// ---- DUTs/IO/Topology/Device_4_EtherCAT_07442C6B.TcDUT
{attribute 'GeneratedUsingTerminal: IODEVICETYPE_ETHERCATPROT'}
{attribute addProperty BoxType "IODEVICETYPE_ETHERCATPROT"}
{attribute addProperty Id "R1_EK1100R1_EK1100_4AD22B7B1143R2_EK1100R2_EK1100_10D8A594458R3_EK1100R3_EK1100_C7887D6C263R4_EK1100R4_EK1100_46A1248C369R4A_EK1100R4A_EK1100_48316913274R5_EK1100R5_EK1100_0007A337146R6_EK1100R6_EK1100_8C41F5F2336R7_EK1100R7_EK1100_F50DDAC8306R8_EK1100R8_EK1100_9C7B3B675648R9_EK1100R9_EK1100_484053C0136R10_EK1100R10_EK1100_C5CE1D87649SyncUnitsSyncUnits_5BE71B8B288InputsInputs_A65FACA410OutputsOutputs_23C0ED1D6InfoDataInfoData_84133AC922"}
{attribute addProperty CRC "121908331"}
{attribute addProperty Size "10054"}
{attribute addProperty Name "Device 4 (EtherCAT)"}
TYPE Device_4_EtherCAT_07442C6B EXTENDS TcoIo.EtcMasterBase_62654B43 :
STRUCT
	{attribute addProperty Name "R1 (EK1100)"}
	{attribute addProperty PreviousPort "Device 4 (EtherCAT) : Master"}
	{attribute addProperty SyncUnit "default"}
	R1_EK1100 : R1_EK1100_4AD22B7B;
	{attribute addProperty Name "R2 (EK1100)"}
	{attribute addProperty PreviousPort "R1 (EK1100) : C"}
	{attribute addProperty SyncUnit "default"}
	R2_EK1100 : R2_EK1100_10D8A594;
	{attribute addProperty Name "R3 (EK1100)"}
	{attribute addProperty PreviousPort "R2 (EK1100) : C"}
	{attribute addProperty SyncUnit "default"}
	R3_EK1100 : R3_EK1100_C7887D6C;
	{attribute addProperty Name "R4 (EK1100)"}
	{attribute addProperty PreviousPort "R3 (EK1100) : C"}
	{attribute addProperty SyncUnit "default"}
	R4_EK1100 : R4_EK1100_46A1248C;
	{attribute addProperty Name "R4A (EK1100)"}
	{attribute addProperty PreviousPort "R4 (EK1100) : C"}
	{attribute addProperty SyncUnit "default"}
	R4A_EK1100 : R4A_EK1100_48316913;
	{attribute addProperty Name "R5 (EK1100)"}
	{attribute addProperty PreviousPort "R4A (EK1100) : C"}
	{attribute addProperty SyncUnit "default"}
	R5_EK1100 : R5_EK1100_0007A337;
	{attribute addProperty Name "R6 (EK1100)"}
	{attribute addProperty PreviousPort "R5 (EK1100) : C"}
	{attribute addProperty SyncUnit "default"}
	R6_EK1100 : R6_EK1100_8C41F5F2;
	{attribute addProperty Name "R7 (EK1100)"}
	{attribute addProperty PreviousPort "R6 (EK1100) : C"}
	{attribute addProperty SyncUnit "default"}
	R7_EK1100 : R7_EK1100_F50DDAC8;
	{attribute addProperty Name "R8 (EK1100)"}
	{attribute addProperty PreviousPort "R7 (EK1100) : C"}
	{attribute addProperty SyncUnit "default"}
	R8_EK1100 : R8_EK1100_9C7B3B67;
	{attribute addProperty Name "R9 (EK1100)"}
	{attribute addProperty PreviousPort "R8 (EK1100) : C"}
	{attribute addProperty SyncUnit "default"}
	R9_EK1100 : R9_EK1100_484053C0;
	{attribute addProperty Name "R10 (EK1100)"}
	{attribute addProperty PreviousPort "R9 (EK1100) : C"}
	{attribute addProperty SyncUnit "default"}
	R10_EK1100 : R10_EK1100_C5CE1D87;
	{attribute addProperty Name "SyncUnits"}
	SyncUnits : SyncUnits_5BE71B8B;
	{attribute addProperty Name "Inputs"}
	Inputs : TcoIo.Inputs_A65FACA4;
	{attribute addProperty Name "Outputs"}
	Outputs : TcoIo.Outputs_23C0ED1D;
	{attribute addProperty Name "InfoData"}
	InfoData : TcoIo.InfoData_84133AC9;
END_STRUCT
END_TYPE

// ---- DUTs/IO/Topology/Term_279_EK1100_ED7D6272.TcDUT
{attribute 'GeneratedUsingTerminal: EK1100-0000-0018'}
{attribute addProperty BoxType "EK1100-0000-0018"}
{attribute addProperty Id "Term_280_EL1809EL1809_32157CFD20Term_281_EL1809EL1809_32157CFD20Term_282_EL1809EL1809_32157CFD20Term_283_EL1809EL1809_32157CFD20Term_284_EL1809EL1809_32157CFD20Term_312_EL1809EL1809_32157CFD20Term_320_EL1809EL1809_32157CFD20Term_321_EL1809EL1809_32157CFD20Term_322_EL1809EL1809_32157CFD20Term_323_EL1809EL1809_32157CFD20Term_324_EL1809EL1809_32157CFD20Term_325_EL1809EL1809_32157CFD20Term_326_EL1809EL1809_32157CFD20Term_327_EL1809EL1809_32157CFD20Term_328_EL1809EL1809_32157CFD20Term_329_EL1809EL1809_32157CFD20Term_331_EL1809EL1809_32157CFD20Term_332_EL1809EL1809_32157CFD20Term_333_EL1809EL1809_32157CFD20Term_334_EL1809EL1809_32157CFD20Term_335_EL1809EL1809_32157CFD20Term_336_EL1809EL1809_32157CFD20Term_337_EL1809EL1809_32157CFD20Term_338_EL1809EL1809_32157CFD20Term_339_EL1809EL1809_32157CFD20Term_340_EL1809EL1809_32157CFD20Term_341_EL1809EL1809_32157CFD20Term_342_EL1809EL1809_32157CFD20Term_343_EL1809EL1809_32157CFD20Term_344_EL1809EL1809_32157CFD20Term_345_EL1809EL1809_32157CFD20Term_346_EL1809EL1809_32157CFD20Term_347_EL1809EL1809_32157CFD20Term_348_EL1809EL1809_32157CFD20Term_360_EL1809EL1809_32157CFD20Term_361_EL1809EL1809_32157CFD20Term_362_EL1809EL1809_32157CFD20Term_363_EL1809EL1809_32157CFD20Term_364_EL1809EL1809_32157CFD20Term_365_EL1809EL1809_32157CFD20Term_366_EL1809EL1809_32157CFD20Term_367_EL1809EL1809_32157CFD20Term_368_EL1809EL1809_32157CFD20Term_370_EL1809EL1809_32157CFD20Term_371_EL1809EL1809_32157CFD20Term_372_EL1809EL1809_32157CFD20Term_373_EL1809EL1809_32157CFD20Term_374_EL1809EL1809_32157CFD20Term_375_EL1809EL1809_32157CFD20Term_376_EL1809EL1809_32157CFD20Term_377_EL1809EL1809_32157CFD20Term_378_EL1809EL1809_32157CFD20Term_380_EL1809EL1809_32157CFD20Term_381_EL1809EL1809_32157CFD20Term_382_EL1809EL1809_32157CFD20Term_383_EL1809EL1809_32157CFD20Term_384_EL1809EL1809_32157CFD20Term_385_EL1809EL1809_32157CFD20Term_386_EL1809EL1809_32157CFD20Term_387_EL1809EL1809_32157CFD20Term_388_EL1809EL1809_32157CFD20Term_389_EL1809EL1809_32157CFD20Term_390_EL1809EL1809_32157CFD20Term_391_EL1809EL1809_32157CFD20Term_392_EL1809EL1809_32157CFD20Term_393_EL1809EL1809_32157CFD20Term_394_EL1809EL1809_32157CFD20Term_395_EL1809EL1809_32157CFD20Term_396_EL1809EL1809_32157CFD20Term_397_EL1809EL1809_32157CFD20Term_398_EL1809EL1809_32157CFD20Term_399_EL1809EL1809_32157CFD20Term_400_EL1809EL1809_32157CFD20Term_401_EL1809EL1809_32157CFD20Term_402_EL1809EL1809_32157CFD20Term_403_EL1809EL1809_32157CFD20Term_404_EL1809EL1809_32157CFD20Term_405_EL1809EL1809_32157CFD20Term_406_EL1809EL1809_32157CFD20Term_407_EL1809EL1809_32157CFD20Term_408_EL1809EL1809_32157CFD20Term_409_EL1809EL1809_32157CFD20Term_410_EL1809EL1809_32157CFD20Term_414_EL1809EL1809_32157CFD20Term_415_EL1809EL1809_32157CFD20Term_416_EL1809EL1809_32157CFD20Term_417_EL1809EL1809_32157CFD20Term_418_EL1809EL1809_32157CFD20Term_419_EL1809EL1809_32157CFD20Term_420_EL1809EL1809_32157CFD20Term_421_EL1809EL1809_32157CFD20Term_422_EL1809EL1809_32157CFD20Term_423_EL1809EL1809_32157CFD20Term_424_EL1809EL1809_32157CFD20Term_425_EL1809EL1809_32157CFD20Term_426_EL1809EL1809_32157CFD20Term_427_EL1809EL1809_32157CFD20Term_428_EL1809EL1809_32157CFD20Term_429_EL1809EL1809_32157CFD20Term_448_EL1809EL1809_32157CFD20Term_495_EK1110EK1110_1FC0878B2"}
{attribute addProperty CRC "3984417394"}
{attribute addProperty Size "2002"}
{attribute addProperty Name "Term 279 (EK1100)"}
TYPE Term_279_EK1100_ED7D6272 EXTENDS EK1100_1FC0878B :
STRUCT
	{attribute addProperty Name "Term 280 (EL1809)"}
	{attribute addProperty PreviousPort "Term 279 (EK1100) : B"}
	{attribute addProperty SyncUnit "default"}
	Term_280_EL1809 : EL1809_32157CFD;
	{attribute addProperty Name "Term 281 (EL1809)"}
	{attribute addProperty PreviousPort "Term 280 (EL1809) : B"}
	{attribute addProperty SyncUnit "default"}
	Term_281_EL1809 : EL1809_32157CFD;
	{attribute addProperty Name "Term 282 (EL1809)"}
	{attribute addProperty PreviousPort "Term 281 (EL1809) : B"}
	{attribute addProperty SyncUnit "default"}
	Term_282_EL1809 : EL1809_32157CFD;
	{attribute addProperty Name "Term 283 (EL1809)"}
	{attribute addProperty PreviousPort "Term 282 (EL1809) : B"}
	{attribute addProperty SyncUnit "default"}
	Term_283_EL1809 : EL1809_32157CFD;
	{attribute addProperty Name "Term 284 (EL1809)"}
	{attribute addProperty PreviousPort "Term 283 (EL1809) : B"}
	{attribute addProperty SyncUnit "default"}
	Term_284_EL1809 : EL1809_32157CFD;
	{attribute addProperty Name "Term 312 (EL1809)"}
	{attribute addProperty PreviousPort "Term 284 (EL1809) : B"}
	{attribute addProperty SyncUnit "default"}
	Term_312_EL1809 : EL1809_32157CFD;
	{attribute addProperty Name "Term 320 (EL1809)"}
	{attribute addProperty PreviousPort "Term 312 (EL1809) : B"}
	{attribute addProperty SyncUnit "default"}
	Term_320_EL1809 : EL1809_32157CFD;
	{attribute addProperty Name "Term 321 (EL1809)"}
	{attribute addProperty PreviousPort "Term 320 (EL1809) : B"}
	{attribute addProperty SyncUnit "default"}
	Term_321_EL1809 : EL1809_32157CFD;
	{attribute addProperty Name "Term 322 (EL1809)"}
	{attribute addProperty PreviousPort "Term 321 (EL1809) : B"}
	{attribute addProperty SyncUnit "default"}
	Term_322_EL1809 : EL1809_32157CFD;
	{attribute addProperty Name "Term 323 (EL1809)"}
	{attribute addProperty PreviousPort "Term 322 (EL1809) : B"}
	{attribute addProperty SyncUnit "default"}
	Term_323_EL1809 : EL1809_32157CFD;
	{attribute addProperty Name "Term 324 (EL1809)"}
	{attribute addProperty PreviousPort "Term 323 (EL1809) : B"}
	{attribute addProperty SyncUnit "default"}
	Term_324_EL1809 : EL1809_32157CFD;
	{attribute addProperty Name "Term 325 (EL1809)"}
	{attribute addProperty PreviousPort "Term 324 (EL1809) : B"}
	{attribute addProperty SyncUnit "default"}
	Term_325_EL1809 : EL1809_32157CFD;
	{attribute addProperty Name "Term 326 (EL1809)"}
	{attribute addProperty PreviousPort "Term 325 (EL1809) : B"}
	{attribute addProperty SyncUnit "default"}
	Term_326_EL1809 : EL1809_32157CFD;
	{attribute addProperty Name "Term 327 (EL1809)"}
	{attribute addProperty PreviousPort "Term 326 (EL1809) : B"}
	{attribute addProperty SyncUnit "default"}
	Term_327_EL1809 : EL1809_32157CFD;
	{attribute addProperty Name "Term 328 (EL1809)"}
	{attribute addProperty PreviousPort "Term 327 (EL1809) : B"}
	{attribute addProperty SyncUnit "default"}
	Term_328_EL1809 : EL1809_32157CFD;
	{attribute addProperty Name "Term 329 (EL1809)"}
	{attribute addProperty PreviousPort "Term 328 (EL1809) : B"}
	{attribute addProperty SyncUnit "default"}
	Term_329_EL1809 : EL1809_32157CFD;
	{attribute addProperty Name "Term 331 (EL1809)"}
	{attribute addProperty PreviousPort "Term 329 (EL1809) : B"}
	{attribute addProperty SyncUnit "default"}
	Term_331_EL1809 : EL1809_32157CFD;
	{attribute addProperty Name "Term 332 (EL1809)"}
	{attribute addProperty PreviousPort "Term 331 (EL1809) : B"}
	{attribute addProperty SyncUnit "default"}
	Term_332_EL1809 : EL1809_32157CFD;
	{attribute addProperty Name "Term 333 (EL1809)"}
	{attribute addProperty PreviousPort "Term 332 (EL1809) : B"}
	{attribute addProperty SyncUnit "default"}
	Term_333_EL1809 : EL1809_32157CFD;
	{attribute addProperty Name "Term 334 (EL1809)"}
	{attribute addProperty PreviousPort "Term 333 (EL1809) : B"}
	{attribute addProperty SyncUnit "default"}
	Term_334_EL1809 : EL1809_32157CFD;
	{attribute addProperty Name "Term 335 (EL1809)"}
	{attribute addProperty PreviousPort "Term 334 (EL1809) : B"}
	{attribute addProperty SyncUnit "default"}
	Term_335_EL1809 : EL1809_32157CFD;
	{attribute addProperty Name "Term 336 (EL1809)"}
	{attribute addProperty PreviousPort "Term 335 (EL1809) : B"}
	{attribute addProperty SyncUnit "default"}
	Term_336_EL1809 : EL1809_32157CFD;
	{attribute addProperty Name "Term 337 (EL1809)"}
	{attribute addProperty PreviousPort "Term 336 (EL1809) : B"}
	{attribute addProperty SyncUnit "default"}
	Term_337_EL1809 : EL1809_32157CFD;
	{attribute addProperty Name "Term 338 (EL1809)"}
	{attribute addProperty PreviousPort "Term 337 (EL1809) : B"}
	{attribute addProperty SyncUnit "default"}
	Term_338_EL1809 : EL1809_32157CFD;
	{attribute addProperty Name "Term 339 (EL1809)"}
	{attribute addProperty PreviousPort "Term 338 (EL1809) : B"}
	{attribute addProperty SyncUnit "default"}
	Term_339_EL1809 : EL1809_32157CFD;
	{attribute addProperty Name "Term 340 (EL1809)"}
	{attribute addProperty PreviousPort "Term 339 (EL1809) : B"}
	{attribute addProperty SyncUnit "default"}
	Term_340_EL1809 : EL1809_32157CFD;
	{attribute addProperty Name "Term 341 (EL1809)"}
	{attribute addProperty PreviousPort "Term 340 (EL1809) : B"}
	{attribute addProperty SyncUnit "default"}
	Term_341_EL1809 : EL1809_32157CFD;
	{attribute addProperty Name "Term 342 (EL1809)"}
	{attribute addProperty PreviousPort "Term 341 (EL1809) : B"}
	{attribute addProperty SyncUnit "default"}
	Term_342_EL1809 : EL1809_32157CFD;
	{attribute addProperty Name "Term 343 (EL1809)"}
	{attribute addProperty PreviousPort "Term 342 (EL1809) : B"}
	{attribute addProperty SyncUnit "default"}
	Term_343_EL1809 : EL1809_32157CFD;
	{attribute addProperty Name "Term 344 (EL1809)"}
	{attribute addProperty PreviousPort "Term 343 (EL1809) : B"}
	{attribute addProperty SyncUnit "default"}
	Term_344_EL1809 : EL1809_32157CFD;
	{attribute addProperty Name "Term 345 (EL1809)"}
	{attribute addProperty PreviousPort "Term 344 (EL1809) : B"}
	{attribute addProperty SyncUnit "default"}
	Term_345_EL1809 : EL1809_32157CFD;
	{attribute addProperty Name "Term 346 (EL1809)"}
	{attribute addProperty PreviousPort "Term 345 (EL1809) : B"}
	{attribute addProperty SyncUnit "default"}
	Term_346_EL1809 : EL1809_32157CFD;
	{attribute addProperty Name "Term 347 (EL1809)"}
	{attribute addProperty PreviousPort "Term 346 (EL1809) : B"}
	{attribute addProperty SyncUnit "default"}
	Term_347_EL1809 : EL1809_32157CFD;
	{attribute addProperty Name "Term 348 (EL1809)"}
	{attribute addProperty PreviousPort "Term 347 (EL1809) : B"}
	{attribute addProperty SyncUnit "default"}
	Term_348_EL1809 : EL1809_32157CFD;
	{attribute addProperty Name "Term 360 (EL1809)"}
	{attribute addProperty PreviousPort "Term 348 (EL1809) : B"}
	{attribute addProperty SyncUnit "default"}
	Term_360_EL1809 : EL1809_32157CFD;
	{attribute addProperty Name "Term 361 (EL1809)"}
	{attribute addProperty PreviousPort "Term 360 (EL1809) : B"}
	{attribute addProperty SyncUnit "default"}
	Term_361_EL1809 : EL1809_32157CFD;
	{attribute addProperty Name "Term 362 (EL1809)"}
	{attribute addProperty PreviousPort "Term 361 (EL1809) : B"}
	{attribute addProperty SyncUnit "default"}
	Term_362_EL1809 : EL1809_32157CFD;
	{attribute addProperty Name "Term 363 (EL1809)"}
	{attribute addProperty PreviousPort "Term 362 (EL1809) : B"}
	{attribute addProperty SyncUnit "default"}
	Term_363_EL1809 : EL1809_32157CFD;
	{attribute addProperty Name "Term 364 (EL1809)"}
	{attribute addProperty PreviousPort "Term 363 (EL1809) : B"}
	{attribute addProperty SyncUnit "default"}
	Term_364_EL1809 : EL1809_32157CFD;
	{attribute addProperty Name "Term 365 (EL1809)"}
	{attribute addProperty PreviousPort "Term 364 (EL1809) : B"}
	{attribute addProperty SyncUnit "default"}
	Term_365_EL1809 : EL1809_32157CFD;
	{attribute addProperty Name "Term 366 (EL1809)"}
	{attribute addProperty PreviousPort "Term 365 (EL1809) : B"}
	{attribute addProperty SyncUnit "default"}
	Term_366_EL1809 : EL1809_32157CFD;
	{attribute addProperty Name "Term 367 (EL1809)"}
	{attribute addProperty PreviousPort "Term 366 (EL1809) : B"}
	{attribute addProperty SyncUnit "default"}
	Term_367_EL1809 : EL1809_32157CFD;
	{attribute addProperty Name "Term 368 (EL1809)"}
	{attribute addProperty PreviousPort "Term 367 (EL1809) : B"}
	{attribute addProperty SyncUnit "default"}
	Term_368_EL1809 : EL1809_32157CFD;
	{attribute addProperty Name "Term 370 (EL1809)"}
	{attribute addProperty PreviousPort "Term 368 (EL1809) : B"}
	{attribute addProperty SyncUnit "default"}
	Term_370_EL1809 : EL1809_32157CFD;
	{attribute addProperty Name "Term 371 (EL1809)"}
	{attribute addProperty PreviousPort "Term 370 (EL1809) : B"}
	{attribute addProperty SyncUnit "default"}
	Term_371_EL1809 : EL1809_32157CFD;
	{attribute addProperty Name "Term 372 (EL1809)"}
	{attribute addProperty PreviousPort "Term 371 (EL1809) : B"}
	{attribute addProperty SyncUnit "default"}
	Term_372_EL1809 : EL1809_32157CFD;
	{attribute addProperty Name "Term 373 (EL1809)"}
	{attribute addProperty PreviousPort "Term 372 (EL1809) : B"}
	{attribute addProperty SyncUnit "default"}
	Term_373_EL1809 : EL1809_32157CFD;
	{attribute addProperty Name "Term 374 (EL1809)"}
	{attribute addProperty PreviousPort "Term 373 (EL1809) : B"}
	{attribute addProperty SyncUnit "default"}
	Term_374_EL1809 : EL1809_32157CFD;
	{attribute addProperty Name "Term 375 (EL1809)"}
	{attribute addProperty PreviousPort "Term 374 (EL1809) : B"}
	{attribute addProperty SyncUnit "default"}
	Term_375_EL1809 : EL1809_32157CFD;
	{attribute addProperty Name "Term 376 (EL1809)"}
	{attribute addProperty PreviousPort "Term 375 (EL1809) : B"}
	{attribute addProperty SyncUnit "default"}
	Term_376_EL1809 : EL1809_32157CFD;
	{attribute addProperty Name "Term 377 (EL1809)"}
	{attribute addProperty PreviousPort "Term 376 (EL1809) : B"}
	{attribute addProperty SyncUnit "default"}
	Term_377_EL1809 : EL1809_32157CFD;
	{attribute addProperty Name "Term 378 (EL1809)"}
	{attribute addProperty PreviousPort "Term 377 (EL1809) : B"}
	{attribute addProperty SyncUnit "default"}
	Term_378_EL1809 : EL1809_32157CFD;
	{attribute addProperty Name "Term 380 (EL1809)"}
	{attribute addProperty PreviousPort "Term 378 (EL1809) : B"}
	{attribute addProperty SyncUnit "default"}
	Term_380_EL1809 : EL1809_32157CFD;
	{attribute addProperty Name "Term 381 (EL1809)"}
	{attribute addProperty PreviousPort "Term 380 (EL1809) : B"}
	{attribute addProperty SyncUnit "default"}
	Term_381_EL1809 : EL1809_32157CFD;
	{attribute addProperty Name "Term 382 (EL1809)"}
	{attribute addProperty PreviousPort "Term 381 (EL1809) : B"}
	{attribute addProperty SyncUnit "default"}
	Term_382_EL1809 : EL1809_32157CFD;
	{attribute addProperty Name "Term 383 (EL1809)"}
	{attribute addProperty PreviousPort "Term 382 (EL1809) : B"}
	{attribute addProperty SyncUnit "default"}
	Term_383_EL1809 : EL1809_32157CFD;
	{attribute addProperty Name "Term 384 (EL1809)"}
	{attribute addProperty PreviousPort "Term 383 (EL1809) : B"}
	{attribute addProperty SyncUnit "default"}
	Term_384_EL1809 : EL1809_32157CFD;
	{attribute addProperty Name "Term 385 (EL1809)"}
	{attribute addProperty PreviousPort "Term 384 (EL1809) : B"}
	{attribute addProperty SyncUnit "default"}
	Term_385_EL1809 : EL1809_32157CFD;
	{attribute addProperty Name "Term 386 (EL1809)"}
	{attribute addProperty PreviousPort "Term 385 (EL1809) : B"}
	{attribute addProperty SyncUnit "default"}
	Term_386_EL1809 : EL1809_32157CFD;
	{attribute addProperty Name "Term 387 (EL1809)"}
	{attribute addProperty PreviousPort "Term 386 (EL1809) : B"}
	{attribute addProperty SyncUnit "default"}
	Term_387_EL1809 : EL1809_32157CFD;
	{attribute addProperty Name "Term 388 (EL1809)"}
	{attribute addProperty PreviousPort "Term 387 (EL1809) : B"}
	{attribute addProperty SyncUnit "default"}
	Term_388_EL1809 : EL1809_32157CFD;
	{attribute addProperty Name "Term 389 (EL1809)"}
	{attribute addProperty PreviousPort "Term 388 (EL1809) : B"}
	{attribute addProperty SyncUnit "default"}
	Term_389_EL1809 : EL1809_32157CFD;
	{attribute addProperty Name "Term 390 (EL1809)"}
	{attribute addProperty PreviousPort "Term 389 (EL1809) : B"}
	{attribute addProperty SyncUnit "default"}
	Term_390_EL1809 : EL1809_32157CFD;
	{attribute addProperty Name "Term 391 (EL1809)"}
	{attribute addProperty PreviousPort "Term 390 (EL1809) : B"}
	{attribute addProperty SyncUnit "default"}
	Term_391_EL1809 : EL1809_32157CFD;
	{attribute addProperty Name "Term 392 (EL1809)"}
	{attribute addProperty PreviousPort "Term 391 (EL1809) : B"}
	{attribute addProperty SyncUnit "default"}
	Term_392_EL1809 : EL1809_32157CFD;
	{attribute addProperty Name "Term 393 (EL1809)"}
	{attribute addProperty PreviousPort "Term 392 (EL1809) : B"}
	{attribute addProperty SyncUnit "default"}
	Term_393_EL1809 : EL1809_32157CFD;
	{attribute addProperty Name "Term 394 (EL1809)"}
	{attribute addProperty PreviousPort "Term 393 (EL1809) : B"}
	{attribute addProperty SyncUnit "default"}
	Term_394_EL1809 : EL1809_32157CFD;
	{attribute addProperty Name "Term 395 (EL1809)"}
	{attribute addProperty PreviousPort "Term 394 (EL1809) : B"}
	{attribute addProperty SyncUnit "default"}
	Term_395_EL1809 : EL1809_32157CFD;
	{attribute addProperty Name "Term 396 (EL1809)"}
	{attribute addProperty PreviousPort "Term 395 (EL1809) : B"}
	{attribute addProperty SyncUnit "default"}
	Term_396_EL1809 : EL1809_32157CFD;
	{attribute addProperty Name "Term 397 (EL1809)"}
	{attribute addProperty PreviousPort "Term 396 (EL1809) : B"}
	{attribute addProperty SyncUnit "default"}
	Term_397_EL1809 : EL1809_32157CFD;
	{attribute addProperty Name "Term 398 (EL1809)"}
	{attribute addProperty PreviousPort "Term 397 (EL1809) : B"}
	{attribute addProperty SyncUnit "default"}
	Term_398_EL1809 : EL1809_32157CFD;
	{attribute addProperty Name "Term 399 (EL1809)"}
	{attribute addProperty PreviousPort "Term 398 (EL1809) : B"}
	{attribute addProperty SyncUnit "default"}
	Term_399_EL1809 : EL1809_32157CFD;
	{attribute addProperty Name "Term 400 (EL1809)"}
	{attribute addProperty PreviousPort "Term 399 (EL1809) : B"}
	{attribute addProperty SyncUnit "default"}
	Term_400_EL1809 : EL1809_32157CFD;
	{attribute addProperty Name "Term 401 (EL1809)"}
	{attribute addProperty PreviousPort "Term 400 (EL1809) : B"}
	{attribute addProperty SyncUnit "default"}
	Term_401_EL1809 : EL1809_32157CFD;
	{attribute addProperty Name "Term 402 (EL1809)"}
	{attribute addProperty PreviousPort "Term 401 (EL1809) : B"}
	{attribute addProperty SyncUnit "default"}
	Term_402_EL1809 : EL1809_32157CFD;
	{attribute addProperty Name "Term 403 (EL1809)"}
	{attribute addProperty PreviousPort "Term 402 (EL1809) : B"}
	{attribute addProperty SyncUnit "default"}
	Term_403_EL1809 : EL1809_32157CFD;
	{attribute addProperty Name "Term 404 (EL1809)"}
	{attribute addProperty PreviousPort "Term 403 (EL1809) : B"}
	{attribute addProperty SyncUnit "default"}
	Term_404_EL1809 : EL1809_32157CFD;
	{attribute addProperty Name "Term 405 (EL1809)"}
	{attribute addProperty PreviousPort "Term 404 (EL1809) : B"}
	{attribute addProperty SyncUnit "default"}
	Term_405_EL1809 : EL1809_32157CFD;
	{attribute addProperty Name "Term 406 (EL1809)"}
	{attribute addProperty PreviousPort "Term 405 (EL1809) : B"}
	{attribute addProperty SyncUnit "default"}
	Term_406_EL1809 : EL1809_32157CFD;
	{attribute addProperty Name "Term 407 (EL1809)"}
	{attribute addProperty PreviousPort "Term 406 (EL1809) : B"}
	{attribute addProperty SyncUnit "default"}
	Term_407_EL1809 : EL1809_32157CFD;
	{attribute addProperty Name "Term 408 (EL1809)"}
	{attribute addProperty PreviousPort "Term 407 (EL1809) : B"}
	{attribute addProperty SyncUnit "default"}
	Term_408_EL1809 : EL1809_32157CFD;
	{attribute addProperty Name "Term 409 (EL1809)"}
	{attribute addProperty PreviousPort "Term 408 (EL1809) : B"}
	{attribute addProperty SyncUnit "default"}
	Term_409_EL1809 : EL1809_32157CFD;
	{attribute addProperty Name "Term 410 (EL1809)"}
	{attribute addProperty PreviousPort "Term 409 (EL1809) : B"}
	{attribute addProperty SyncUnit "default"}
	Term_410_EL1809 : EL1809_32157CFD;
	{attribute addProperty Name "Term 414 (EL1809)"}
	{attribute addProperty PreviousPort "Term 410 (EL1809) : B"}
	{attribute addProperty SyncUnit "default"}
	Term_414_EL1809 : EL1809_32157CFD;
	{attribute addProperty Name "Term 415 (EL1809)"}
	{attribute addProperty PreviousPort "Term 414 (EL1809) : B"}
	{attribute addProperty SyncUnit "default"}
	Term_415_EL1809 : EL1809_32157CFD;
	{attribute addProperty Name "Term 416 (EL1809)"}
	{attribute addProperty PreviousPort "Term 415 (EL1809) : B"}
	{attribute addProperty SyncUnit "default"}
	Term_416_EL1809 : EL1809_32157CFD;
	{attribute addProperty Name "Term 417 (EL1809)"}
	{attribute addProperty PreviousPort "Term 416 (EL1809) : B"}
	{attribute addProperty SyncUnit "default"}
	Term_417_EL1809 : EL1809_32157CFD;
	{attribute addProperty Name "Term 418 (EL1809)"}
	{attribute addProperty PreviousPort "Term 417 (EL1809) : B"}
	{attribute addProperty SyncUnit "default"}
	Term_418_EL1809 : EL1809_32157CFD;
	{attribute addProperty Name "Term 419 (EL1809)"}
	{attribute addProperty PreviousPort "Term 418 (EL1809) : B"}
	{attribute addProperty SyncUnit "default"}
	Term_419_EL1809 : EL1809_32157CFD;
	{attribute addProperty Name "Term 420 (EL1809)"}
	{attribute addProperty PreviousPort "Term 419 (EL1809) : B"}
	{attribute addProperty SyncUnit "default"}
	Term_420_EL1809 : EL1809_32157CFD;
	{attribute addProperty Name "Term 421 (EL1809)"}
	{attribute addProperty PreviousPort "Term 420 (EL1809) : B"}
	{attribute addProperty SyncUnit "default"}
	Term_421_EL1809 : EL1809_32157CFD;
	{attribute addProperty Name "Term 422 (EL1809)"}
	{attribute addProperty PreviousPort "Term 421 (EL1809) : B"}
	{attribute addProperty SyncUnit "default"}
	Term_422_EL1809 : EL1809_32157CFD;
	{attribute addProperty Name "Term 423 (EL1809)"}
	{attribute addProperty PreviousPort "Term 422 (EL1809) : B"}
	{attribute addProperty SyncUnit "default"}
	Term_423_EL1809 : EL1809_32157CFD;
	{attribute addProperty Name "Term 424 (EL1809)"}
	{attribute addProperty PreviousPort "Term 423 (EL1809) : B"}
	{attribute addProperty SyncUnit "default"}
	Term_424_EL1809 : EL1809_32157CFD;
	{attribute addProperty Name "Term 425 (EL1809)"}
	{attribute addProperty PreviousPort "Term 424 (EL1809) : B"}
	{attribute addProperty SyncUnit "default"}
	Term_425_EL1809 : EL1809_32157CFD;
	{attribute addProperty Name "Term 426 (EL1809)"}
	{attribute addProperty PreviousPort "Term 425 (EL1809) : B"}
	{attribute addProperty SyncUnit "default"}
	Term_426_EL1809 : EL1809_32157CFD;
	{attribute addProperty Name "Term 427 (EL1809)"}
	{attribute addProperty PreviousPort "Term 426 (EL1809) : B"}
	{attribute addProperty SyncUnit "default"}
	Term_427_EL1809 : EL1809_32157CFD;
	{attribute addProperty Name "Term 428 (EL1809)"}
	{attribute addProperty PreviousPort "Term 427 (EL1809) : B"}
	{attribute addProperty SyncUnit "default"}
	Term_428_EL1809 : EL1809_32157CFD;
	{attribute addProperty Name "Term 429 (EL1809)"}
	{attribute addProperty PreviousPort "Term 428 (EL1809) : B"}
	{attribute addProperty SyncUnit "default"}
	Term_429_EL1809 : EL1809_32157CFD;
	{attribute addProperty Name "Term 448 (EL1809)"}
	{attribute addProperty PreviousPort "Term 429 (EL1809) : B"}
	{attribute addProperty SyncUnit "default"}
	Term_448_EL1809 : EL1809_32157CFD;
	{attribute addProperty Name "Term 495 (EK1110)"}
	{attribute addProperty PreviousPort "Term 448 (EL1809) : B"}
	{attribute addProperty SyncUnit "default"}
	Term_495_EK1110 : EK1110_1FC0878B;
END_STRUCT
END_TYPE

// ---- DUTs/IO/Topology/Term_554_EK1100_B580E218.TcDUT
{attribute 'GeneratedUsingTerminal: EK1100-0000-0018'}
{attribute addProperty BoxType "EK1100-0000-0018"}
{attribute addProperty Id "Term_645_EL1809EL1809_32157CFD20Term_646_EL1809EL1809_32157CFD20Term_647_EL1809EL1809_32157CFD20Term_648_EL1809EL1809_32157CFD20Term_649_EL1809EL1809_32157CFD20Term_650_EL1809EL1809_32157CFD20Term_651_EL1809EL1809_32157CFD20Term_652_EL1809EL1809_32157CFD20Term_653_EL1809EL1809_32157CFD20Term_654_EL1809EL1809_32157CFD20Term_655_EL1809EL1809_32157CFD20Term_656_EL1809EL1809_32157CFD20Term_657_EL1809EL1809_32157CFD20Term_658_EL1809EL1809_32157CFD20Term_659_EL1809EL1809_32157CFD20Term_660_EL1809EL1809_32157CFD20Term_661_EL1809EL1809_32157CFD20Term_662_EL1809EL1809_32157CFD20Term_663_EL1809EL1809_32157CFD20Term_664_EL1809EL1809_32157CFD20Term_665_EL1809EL1809_32157CFD20Term_666_EL1809EL1809_32157CFD20Term_667_EL1809EL1809_32157CFD20Term_668_EL1809EL1809_32157CFD20Term_669_EL1809EL1809_32157CFD20Term_670_EL1809EL1809_32157CFD20Term_671_EL1809EL1809_32157CFD20Term_672_EL1809EL1809_32157CFD20Term_673_EL1809EL1809_32157CFD20Term_674_EL1809EL1809_32157CFD20Term_676_EL1809EL1809_32157CFD20Term_677_EL1809EL1809_32157CFD20Term_678_EL1809EL1809_32157CFD20Term_679_EL1809EL1809_32157CFD20Term_680_EL1809EL1809_32157CFD20Term_681_EL1809EL1809_32157CFD20Term_682_EL1809EL1809_32157CFD20Term_683_EL1809EL1809_32157CFD20Term_684_EL1809EL1809_32157CFD20Term_685_EL1809EL1809_32157CFD20Term_686_EL1809EL1809_32157CFD20Term_687_EL1809EL1809_32157CFD20Term_688_EL1809EL1809_32157CFD20Term_689_EL1809EL1809_32157CFD20Term_690_EL1809EL1809_32157CFD20Term_691_EL1809EL1809_32157CFD20Term_692_EL1809EL1809_32157CFD20Term_693_EL1809EL1809_32157CFD20Term_694_EL1809EL1809_32157CFD20Term_695_EL1809EL1809_32157CFD20Term_696_EL1809EL1809_32157CFD20Term_697_EL1809EL1809_32157CFD20Term_698_EL1809EL1809_32157CFD20Term_699_EL1809EL1809_32157CFD20Term_700_EL1809EL1809_32157CFD20Term_701_EL1809EL1809_32157CFD20Term_702_EL1809EL1809_32157CFD20Term_703_EL1809EL1809_32157CFD20Term_704_EL1809EL1809_32157CFD20Term_705_EL1809EL1809_32157CFD20Term_706_EL1809EL1809_32157CFD20Term_707_EL1809EL1809_32157CFD20Term_709_EL1809EL1809_32157CFD20Term_710_EL1809EL1809_32157CFD20Term_711_EL1809EL1809_32157CFD20Term_712_EL1809EL1809_32157CFD20Term_713_EL1809EL1809_32157CFD20Term_714_EL1809EL1809_32157CFD20Term_715_EL1809EL1809_32157CFD20Term_716_EL1809EL1809_32157CFD20Term_717_EL1809EL1809_32157CFD20Term_718_EL1809EL1809_32157CFD20Term_719_EL1809EL1809_32157CFD20Term_720_EL1809EL1809_32157CFD20Term_721_EL1809EL1809_32157CFD20Term_722_EL1809EL1809_32157CFD20Term_723_EL1809EL1809_32157CFD20Term_724_EL1809EL1809_32157CFD20Term_725_EL1809EL1809_32157CFD20Term_726_EL1809EL1809_32157CFD20Term_727_EL1809EL1809_32157CFD20Term_728_EL1809EL1809_32157CFD20Term_729_EL1809EL1809_32157CFD20Term_730_EL1809EL1809_32157CFD20Term_731_EL1809EL1809_32157CFD20Term_732_EL1809EL1809_32157CFD20Term_733_EL1809EL1809_32157CFD20Term_734_EL1809EL1809_32157CFD20Term_735_EL1809EL1809_32157CFD20Term_736_EL1809EL1809_32157CFD20Term_737_EL1809EL1809_32157CFD20Term_738_EL1809EL1809_32157CFD20Term_739_EL1809EL1809_32157CFD20Term_740_EL1809EL1809_32157CFD20Term_741_EL1809EL1809_32157CFD20Term_742_EL1809EL1809_32157CFD20Term_743_EL1809EL1809_32157CFD20Term_744_EL1809EL1809_32157CFD20Term_745_EL1809EL1809_32157CFD20Term_746_EL1809EL1809_32157CFD20Term_747_EK1110EK1110_1FC0878B2"}
{attribute addProperty CRC "3045122584"}
{attribute addProperty Size "2002"}
{attribute addProperty Name "Term 554 (EK1100)"}
TYPE Term_554_EK1100_B580E218 EXTENDS EK1100_1FC0878B :
STRUCT
	{attribute addProperty Name "Term 645 (EL1809)"}
	{attribute addProperty PreviousPort "Term 554 (EK1100) : B"}
	{attribute addProperty SyncUnit "default"}
	Term_645_EL1809 : EL1809_32157CFD;
	{attribute addProperty Name "Term 646 (EL1809)"}
	{attribute addProperty PreviousPort "Term 645 (EL1809) : B"}
	{attribute addProperty SyncUnit "default"}
	Term_646_EL1809 : EL1809_32157CFD;
	{attribute addProperty Name "Term 647 (EL1809)"}
	{attribute addProperty PreviousPort "Term 646 (EL1809) : B"}
	{attribute addProperty SyncUnit "default"}
	Term_647_EL1809 : EL1809_32157CFD;
	{attribute addProperty Name "Term 648 (EL1809)"}
	{attribute addProperty PreviousPort "Term 647 (EL1809) : B"}
	{attribute addProperty SyncUnit "default"}
	Term_648_EL1809 : EL1809_32157CFD;
	{attribute addProperty Name "Term 649 (EL1809)"}
	{attribute addProperty PreviousPort "Term 648 (EL1809) : B"}
	{attribute addProperty SyncUnit "default"}
	Term_649_EL1809 : EL1809_32157CFD;
	{attribute addProperty Name "Term 650 (EL1809)"}
	{attribute addProperty PreviousPort "Term 649 (EL1809) : B"}
	{attribute addProperty SyncUnit "default"}
	Term_650_EL1809 : EL1809_32157CFD;
	{attribute addProperty Name "Term 651 (EL1809)"}
	{attribute addProperty PreviousPort "Term 650 (EL1809) : B"}
	{attribute addProperty SyncUnit "default"}
	Term_651_EL1809 : EL1809_32157CFD;
	{attribute addProperty Name "Term 652 (EL1809)"}
	{attribute addProperty PreviousPort "Term 651 (EL1809) : B"}
	{attribute addProperty SyncUnit "default"}
	Term_652_EL1809 : EL1809_32157CFD;
	{attribute addProperty Name "Term 653 (EL1809)"}
	{attribute addProperty PreviousPort "Term 652 (EL1809) : B"}
	{attribute addProperty SyncUnit "default"}
	Term_653_EL1809 : EL1809_32157CFD;
	{attribute addProperty Name "Term 654 (EL1809)"}
	{attribute addProperty PreviousPort "Term 653 (EL1809) : B"}
	{attribute addProperty SyncUnit "default"}
	Term_654_EL1809 : EL1809_32157CFD;
	{attribute addProperty Name "Term 655 (EL1809)"}
	{attribute addProperty PreviousPort "Term 654 (EL1809) : B"}
	{attribute addProperty SyncUnit "default"}
	Term_655_EL1809 : EL1809_32157CFD;
	{attribute addProperty Name "Term 656 (EL1809)"}
	{attribute addProperty PreviousPort "Term 655 (EL1809) : B"}
	{attribute addProperty SyncUnit "default"}
	Term_656_EL1809 : EL1809_32157CFD;
	{attribute addProperty Name "Term 657 (EL1809)"}
	{attribute addProperty PreviousPort "Term 656 (EL1809) : B"}
	{attribute addProperty SyncUnit "default"}
	Term_657_EL1809 : EL1809_32157CFD;
	{attribute addProperty Name "Term 658 (EL1809)"}
	{attribute addProperty PreviousPort "Term 657 (EL1809) : B"}
	{attribute addProperty SyncUnit "default"}
	Term_658_EL1809 : EL1809_32157CFD;
	{attribute addProperty Name "Term 659 (EL1809)"}
	{attribute addProperty PreviousPort "Term 658 (EL1809) : B"}
	{attribute addProperty SyncUnit "default"}
	Term_659_EL1809 : EL1809_32157CFD;
	{attribute addProperty Name "Term 660 (EL1809)"}
	{attribute addProperty PreviousPort "Term 659 (EL1809) : B"}
	{attribute addProperty SyncUnit "default"}
	Term_660_EL1809 : EL1809_32157CFD;
	{attribute addProperty Name "Term 661 (EL1809)"}
	{attribute addProperty PreviousPort "Term 660 (EL1809) : B"}
	{attribute addProperty SyncUnit "default"}
	Term_661_EL1809 : EL1809_32157CFD;
	{attribute addProperty Name "Term 662 (EL1809)"}
	{attribute addProperty PreviousPort "Term 661 (EL1809) : B"}
	{attribute addProperty SyncUnit "default"}
	Term_662_EL1809 : EL1809_32157CFD;
	{attribute addProperty Name "Term 663 (EL1809)"}
	{attribute addProperty PreviousPort "Term 662 (EL1809) : B"}
	{attribute addProperty SyncUnit "default"}
	Term_663_EL1809 : EL1809_32157CFD;
	{attribute addProperty Name "Term 664 (EL1809)"}
	{attribute addProperty PreviousPort "Term 663 (EL1809) : B"}
	{attribute addProperty SyncUnit "default"}
	Term_664_EL1809 : EL1809_32157CFD;
	{attribute addProperty Name "Term 665 (EL1809)"}
	{attribute addProperty PreviousPort "Term 664 (EL1809) : B"}
	{attribute addProperty SyncUnit "default"}
	Term_665_EL1809 : EL1809_32157CFD;
	{attribute addProperty Name "Term 666 (EL1809)"}
	{attribute addProperty PreviousPort "Term 665 (EL1809) : B"}
	{attribute addProperty SyncUnit "default"}
	Term_666_EL1809 : EL1809_32157CFD;
	{attribute addProperty Name "Term 667 (EL1809)"}
	{attribute addProperty PreviousPort "Term 666 (EL1809) : B"}
	{attribute addProperty SyncUnit "default"}
	Term_667_EL1809 : EL1809_32157CFD;
	{attribute addProperty Name "Term 668 (EL1809)"}
	{attribute addProperty PreviousPort "Term 667 (EL1809) : B"}
	{attribute addProperty SyncUnit "default"}
	Term_668_EL1809 : EL1809_32157CFD;
	{attribute addProperty Name "Term 669 (EL1809)"}
	{attribute addProperty PreviousPort "Term 668 (EL1809) : B"}
	{attribute addProperty SyncUnit "default"}
	Term_669_EL1809 : EL1809_32157CFD;
	{attribute addProperty Name "Term 670 (EL1809)"}
	{attribute addProperty PreviousPort "Term 669 (EL1809) : B"}
	{attribute addProperty SyncUnit "default"}
	Term_670_EL1809 : EL1809_32157CFD;
	{attribute addProperty Name "Term 671 (EL1809)"}
	{attribute addProperty PreviousPort "Term 670 (EL1809) : B"}
	{attribute addProperty SyncUnit "default"}
	Term_671_EL1809 : EL1809_32157CFD;
	{attribute addProperty Name "Term 672 (EL1809)"}
	{attribute addProperty PreviousPort "Term 671 (EL1809) : B"}
	{attribute addProperty SyncUnit "default"}
	Term_672_EL1809 : EL1809_32157CFD;
	{attribute addProperty Name "Term 673 (EL1809)"}
	{attribute addProperty PreviousPort "Term 672 (EL1809) : B"}
	{attribute addProperty SyncUnit "default"}
	Term_673_EL1809 : EL1809_32157CFD;
	{attribute addProperty Name "Term 674 (EL1809)"}
	{attribute addProperty PreviousPort "Term 673 (EL1809) : B"}
	{attribute addProperty SyncUnit "default"}
	Term_674_EL1809 : EL1809_32157CFD;
	{attribute addProperty Name "Term 676 (EL1809)"}
	{attribute addProperty PreviousPort "Term 674 (EL1809) : B"}
	{attribute addProperty SyncUnit "default"}
	Term_676_EL1809 : EL1809_32157CFD;
	{attribute addProperty Name "Term 677 (EL1809)"}
	{attribute addProperty PreviousPort "Term 676 (EL1809) : B"}
	{attribute addProperty SyncUnit "default"}
	Term_677_EL1809 : EL1809_32157CFD;
	{attribute addProperty Name "Term 678 (EL1809)"}
	{attribute addProperty PreviousPort "Term 677 (EL1809) : B"}
	{attribute addProperty SyncUnit "default"}
	Term_678_EL1809 : EL1809_32157CFD;
	{attribute addProperty Name "Term 679 (EL1809)"}
	{attribute addProperty PreviousPort "Term 678 (EL1809) : B"}
	{attribute addProperty SyncUnit "default"}
	Term_679_EL1809 : EL1809_32157CFD;
	{attribute addProperty Name "Term 680 (EL1809)"}
	{attribute addProperty PreviousPort "Term 679 (EL1809) : B"}
	{attribute addProperty SyncUnit "default"}
	Term_680_EL1809 : EL1809_32157CFD;
	{attribute addProperty Name "Term 681 (EL1809)"}
	{attribute addProperty PreviousPort "Term 680 (EL1809) : B"}
	{attribute addProperty SyncUnit "default"}
	Term_681_EL1809 : EL1809_32157CFD;
	{attribute addProperty Name "Term 682 (EL1809)"}
	{attribute addProperty PreviousPort "Term 681 (EL1809) : B"}
	{attribute addProperty SyncUnit "default"}
	Term_682_EL1809 : EL1809_32157CFD;
	{attribute addProperty Name "Term 683 (EL1809)"}
	{attribute addProperty PreviousPort "Term 682 (EL1809) : B"}
	{attribute addProperty SyncUnit "default"}
	Term_683_EL1809 : EL1809_32157CFD;
	{attribute addProperty Name "Term 684 (EL1809)"}
	{attribute addProperty PreviousPort "Term 683 (EL1809) : B"}
	{attribute addProperty SyncUnit "default"}
	Term_684_EL1809 : EL1809_32157CFD;
	{attribute addProperty Name "Term 685 (EL1809)"}
	{attribute addProperty PreviousPort "Term 684 (EL1809) : B"}
	{attribute addProperty SyncUnit "default"}
	Term_685_EL1809 : EL1809_32157CFD;
	{attribute addProperty Name "Term 686 (EL1809)"}
	{attribute addProperty PreviousPort "Term 685 (EL1809) : B"}
	{attribute addProperty SyncUnit "default"}
	Term_686_EL1809 : EL1809_32157CFD;
	{attribute addProperty Name "Term 687 (EL1809)"}
	{attribute addProperty PreviousPort "Term 686 (EL1809) : B"}
	{attribute addProperty SyncUnit "default"}
	Term_687_EL1809 : EL1809_32157CFD;
	{attribute addProperty Name "Term 688 (EL1809)"}
	{attribute addProperty PreviousPort "Term 687 (EL1809) : B"}
	{attribute addProperty SyncUnit "default"}
	Term_688_EL1809 : EL1809_32157CFD;
	{attribute addProperty Name "Term 689 (EL1809)"}
	{attribute addProperty PreviousPort "Term 688 (EL1809) : B"}
	{attribute addProperty SyncUnit "default"}
	Term_689_EL1809 : EL1809_32157CFD;
	{attribute addProperty Name "Term 690 (EL1809)"}
	{attribute addProperty PreviousPort "Term 689 (EL1809) : B"}
	{attribute addProperty SyncUnit "default"}
	Term_690_EL1809 : EL1809_32157CFD;
	{attribute addProperty Name "Term 691 (EL1809)"}
	{attribute addProperty PreviousPort "Term 690 (EL1809) : B"}
	{attribute addProperty SyncUnit "default"}
	Term_691_EL1809 : EL1809_32157CFD;
	{attribute addProperty Name "Term 692 (EL1809)"}
	{attribute addProperty PreviousPort "Term 691 (EL1809) : B"}
	{attribute addProperty SyncUnit "default"}
	Term_692_EL1809 : EL1809_32157CFD;
	{attribute addProperty Name "Term 693 (EL1809)"}
	{attribute addProperty PreviousPort "Term 692 (EL1809) : B"}
	{attribute addProperty SyncUnit "default"}
	Term_693_EL1809 : EL1809_32157CFD;
	{attribute addProperty Name "Term 694 (EL1809)"}
	{attribute addProperty PreviousPort "Term 693 (EL1809) : B"}
	{attribute addProperty SyncUnit "default"}
	Term_694_EL1809 : EL1809_32157CFD;
	{attribute addProperty Name "Term 695 (EL1809)"}
	{attribute addProperty PreviousPort "Term 694 (EL1809) : B"}
	{attribute addProperty SyncUnit "default"}
	Term_695_EL1809 : EL1809_32157CFD;
	{attribute addProperty Name "Term 696 (EL1809)"}
	{attribute addProperty PreviousPort "Term 695 (EL1809) : B"}
	{attribute addProperty SyncUnit "default"}
	Term_696_EL1809 : EL1809_32157CFD;
	{attribute addProperty Name "Term 697 (EL1809)"}
	{attribute addProperty PreviousPort "Term 696 (EL1809) : B"}
	{attribute addProperty SyncUnit "default"}
	Term_697_EL1809 : EL1809_32157CFD;
	{attribute addProperty Name "Term 698 (EL1809)"}
	{attribute addProperty PreviousPort "Term 697 (EL1809) : B"}
	{attribute addProperty SyncUnit "default"}
	Term_698_EL1809 : EL1809_32157CFD;
	{attribute addProperty Name "Term 699 (EL1809)"}
	{attribute addProperty PreviousPort "Term 698 (EL1809) : B"}
	{attribute addProperty SyncUnit "default"}
	Term_699_EL1809 : EL1809_32157CFD;
	{attribute addProperty Name "Term 700 (EL1809)"}
	{attribute addProperty PreviousPort "Term 699 (EL1809) : B"}
	{attribute addProperty SyncUnit "default"}
	Term_700_EL1809 : EL1809_32157CFD;
	{attribute addProperty Name "Term 701 (EL1809)"}
	{attribute addProperty PreviousPort "Term 700 (EL1809) : B"}
	{attribute addProperty SyncUnit "default"}
	Term_701_EL1809 : EL1809_32157CFD;
	{attribute addProperty Name "Term 702 (EL1809)"}
	{attribute addProperty PreviousPort "Term 701 (EL1809) : B"}
	{attribute addProperty SyncUnit "default"}
	Term_702_EL1809 : EL1809_32157CFD;
	{attribute addProperty Name "Term 703 (EL1809)"}
	{attribute addProperty PreviousPort "Term 702 (EL1809) : B"}
	{attribute addProperty SyncUnit "default"}
	Term_703_EL1809 : EL1809_32157CFD;
	{attribute addProperty Name "Term 704 (EL1809)"}
	{attribute addProperty PreviousPort "Term 703 (EL1809) : B"}
	{attribute addProperty SyncUnit "default"}
	Term_704_EL1809 : EL1809_32157CFD;
	{attribute addProperty Name "Term 705 (EL1809)"}
	{attribute addProperty PreviousPort "Term 704 (EL1809) : B"}
	{attribute addProperty SyncUnit "default"}
	Term_705_EL1809 : EL1809_32157CFD;
	{attribute addProperty Name "Term 706 (EL1809)"}
	{attribute addProperty PreviousPort "Term 705 (EL1809) : B"}
	{attribute addProperty SyncUnit "default"}
	Term_706_EL1809 : EL1809_32157CFD;
	{attribute addProperty Name "Term 707 (EL1809)"}
	{attribute addProperty PreviousPort "Term 706 (EL1809) : B"}
	{attribute addProperty SyncUnit "default"}
	Term_707_EL1809 : EL1809_32157CFD;
	{attribute addProperty Name "Term 709 (EL1809)"}
	{attribute addProperty PreviousPort "Term 707 (EL1809) : B"}
	{attribute addProperty SyncUnit "default"}
	Term_709_EL1809 : EL1809_32157CFD;
	{attribute addProperty Name "Term 710 (EL1809)"}
	{attribute addProperty PreviousPort "Term 709 (EL1809) : B"}
	{attribute addProperty SyncUnit "default"}
	Term_710_EL1809 : EL1809_32157CFD;
	{attribute addProperty Name "Term 711 (EL1809)"}
	{attribute addProperty PreviousPort "Term 710 (EL1809) : B"}
	{attribute addProperty SyncUnit "default"}
	Term_711_EL1809 : EL1809_32157CFD;
	{attribute addProperty Name "Term 712 (EL1809)"}
	{attribute addProperty PreviousPort "Term 711 (EL1809) : B"}
	{attribute addProperty SyncUnit "default"}
	Term_712_EL1809 : EL1809_32157CFD;
	{attribute addProperty Name "Term 713 (EL1809)"}
	{attribute addProperty PreviousPort "Term 712 (EL1809) : B"}
	{attribute addProperty SyncUnit "default"}
	Term_713_EL1809 : EL1809_32157CFD;
	{attribute addProperty Name "Term 714 (EL1809)"}
	{attribute addProperty PreviousPort "Term 713 (EL1809) : B"}
	{attribute addProperty SyncUnit "default"}
	Term_714_EL1809 : EL1809_32157CFD;
	{attribute addProperty Name "Term 715 (EL1809)"}
	{attribute addProperty PreviousPort "Term 714 (EL1809) : B"}
	{attribute addProperty SyncUnit "default"}
	Term_715_EL1809 : EL1809_32157CFD;
	{attribute addProperty Name "Term 716 (EL1809)"}
	{attribute addProperty PreviousPort "Term 715 (EL1809) : B"}
	{attribute addProperty SyncUnit "default"}
	Term_716_EL1809 : EL1809_32157CFD;
	{attribute addProperty Name "Term 717 (EL1809)"}
	{attribute addProperty PreviousPort "Term 716 (EL1809) : B"}
	{attribute addProperty SyncUnit "default"}
	Term_717_EL1809 : EL1809_32157CFD;
	{attribute addProperty Name "Term 718 (EL1809)"}
	{attribute addProperty PreviousPort "Term 717 (EL1809) : B"}
	{attribute addProperty SyncUnit "default"}
	Term_718_EL1809 : EL1809_32157CFD;
	{attribute addProperty Name "Term 719 (EL1809)"}
	{attribute addProperty PreviousPort "Term 718 (EL1809) : B"}
	{attribute addProperty SyncUnit "default"}
	Term_719_EL1809 : EL1809_32157CFD;
	{attribute addProperty Name "Term 720 (EL1809)"}
	{attribute addProperty PreviousPort "Term 719 (EL1809) : B"}
	{attribute addProperty SyncUnit "default"}
	Term_720_EL1809 : EL1809_32157CFD;
	{attribute addProperty Name "Term 721 (EL1809)"}
	{attribute addProperty PreviousPort "Term 720 (EL1809) : B"}
	{attribute addProperty SyncUnit "default"}
	Term_721_EL1809 : EL1809_32157CFD;
	{attribute addProperty Name "Term 722 (EL1809)"}
	{attribute addProperty PreviousPort "Term 721 (EL1809) : B"}
	{attribute addProperty SyncUnit "default"}
	Term_722_EL1809 : EL1809_32157CFD;
	{attribute addProperty Name "Term 723 (EL1809)"}
	{attribute addProperty PreviousPort "Term 722 (EL1809) : B"}
	{attribute addProperty SyncUnit "default"}
	Term_723_EL1809 : EL1809_32157CFD;
	{attribute addProperty Name "Term 724 (EL1809)"}
	{attribute addProperty PreviousPort "Term 723 (EL1809) : B"}
	{attribute addProperty SyncUnit "default"}
	Term_724_EL1809 : EL1809_32157CFD;
	{attribute addProperty Name "Term 725 (EL1809)"}
	{attribute addProperty PreviousPort "Term 724 (EL1809) : B"}
	{attribute addProperty SyncUnit "default"}
	Term_725_EL1809 : EL1809_32157CFD;
	{attribute addProperty Name "Term 726 (EL1809)"}
	{attribute addProperty PreviousPort "Term 725 (EL1809) : B"}
	{attribute addProperty SyncUnit "default"}
	Term_726_EL1809 : EL1809_32157CFD;
	{attribute addProperty Name "Term 727 (EL1809)"}
	{attribute addProperty PreviousPort "Term 726 (EL1809) : B"}
	{attribute addProperty SyncUnit "default"}
	Term_727_EL1809 : EL1809_32157CFD;
	{attribute addProperty Name "Term 728 (EL1809)"}
	{attribute addProperty PreviousPort "Term 727 (EL1809) : B"}
	{attribute addProperty SyncUnit "default"}
	Term_728_EL1809 : EL1809_32157CFD;
	{attribute addProperty Name "Term 729 (EL1809)"}
	{attribute addProperty PreviousPort "Term 728 (EL1809) : B"}
	{attribute addProperty SyncUnit "default"}
	Term_729_EL1809 : EL1809_32157CFD;
	{attribute addProperty Name "Term 730 (EL1809)"}
	{attribute addProperty PreviousPort "Term 729 (EL1809) : B"}
	{attribute addProperty SyncUnit "default"}
	Term_730_EL1809 : EL1809_32157CFD;
	{attribute addProperty Name "Term 731 (EL1809)"}
	{attribute addProperty PreviousPort "Term 730 (EL1809) : B"}
	{attribute addProperty SyncUnit "default"}
	Term_731_EL1809 : EL1809_32157CFD;
	{attribute addProperty Name "Term 732 (EL1809)"}
	{attribute addProperty PreviousPort "Term 731 (EL1809) : B"}
	{attribute addProperty SyncUnit "default"}
	Term_732_EL1809 : EL1809_32157CFD;
	{attribute addProperty Name "Term 733 (EL1809)"}
	{attribute addProperty PreviousPort "Term 732 (EL1809) : B"}
	{attribute addProperty SyncUnit "default"}
	Term_733_EL1809 : EL1809_32157CFD;
	{attribute addProperty Name "Term 734 (EL1809)"}
	{attribute addProperty PreviousPort "Term 733 (EL1809) : B"}
	{attribute addProperty SyncUnit "default"}
	Term_734_EL1809 : EL1809_32157CFD;
	{attribute addProperty Name "Term 735 (EL1809)"}
	{attribute addProperty PreviousPort "Term 734 (EL1809) : B"}
	{attribute addProperty SyncUnit "default"}
	Term_735_EL1809 : EL1809_32157CFD;
	{attribute addProperty Name "Term 736 (EL1809)"}
	{attribute addProperty PreviousPort "Term 735 (EL1809) : B"}
	{attribute addProperty SyncUnit "default"}
	Term_736_EL1809 : EL1809_32157CFD;
	{attribute addProperty Name "Term 737 (EL1809)"}
	{attribute addProperty PreviousPort "Term 736 (EL1809) : B"}
	{attribute addProperty SyncUnit "default"}
	Term_737_EL1809 : EL1809_32157CFD;
	{attribute addProperty Name "Term 738 (EL1809)"}
	{attribute addProperty PreviousPort "Term 737 (EL1809) : B"}
	{attribute addProperty SyncUnit "default"}
	Term_738_EL1809 : EL1809_32157CFD;
	{attribute addProperty Name "Term 739 (EL1809)"}
	{attribute addProperty PreviousPort "Term 738 (EL1809) : B"}
	{attribute addProperty SyncUnit "default"}
	Term_739_EL1809 : EL1809_32157CFD;
	{attribute addProperty Name "Term 740 (EL1809)"}
	{attribute addProperty PreviousPort "Term 739 (EL1809) : B"}
	{attribute addProperty SyncUnit "default"}
	Term_740_EL1809 : EL1809_32157CFD;
	{attribute addProperty Name "Term 741 (EL1809)"}
	{attribute addProperty PreviousPort "Term 740 (EL1809) : B"}
	{attribute addProperty SyncUnit "default"}
	Term_741_EL1809 : EL1809_32157CFD;
	{attribute addProperty Name "Term 742 (EL1809)"}
	{attribute addProperty PreviousPort "Term 741 (EL1809) : B"}
	{attribute addProperty SyncUnit "default"}
	Term_742_EL1809 : EL1809_32157CFD;
	{attribute addProperty Name "Term 743 (EL1809)"}
	{attribute addProperty PreviousPort "Term 742 (EL1809) : B"}
	{attribute addProperty SyncUnit "default"}
	Term_743_EL1809 : EL1809_32157CFD;
	{attribute addProperty Name "Term 744 (EL1809)"}
	{attribute addProperty PreviousPort "Term 743 (EL1809) : B"}
	{attribute addProperty SyncUnit "default"}
	Term_744_EL1809 : EL1809_32157CFD;
	{attribute addProperty Name "Term 745 (EL1809)"}
	{attribute addProperty PreviousPort "Term 744 (EL1809) : B"}
	{attribute addProperty SyncUnit "default"}
	Term_745_EL1809 : EL1809_32157CFD;
	{attribute addProperty Name "Term 746 (EL1809)"}
	{attribute addProperty PreviousPort "Term 745 (EL1809) : B"}
	{attribute addProperty SyncUnit "default"}
	Term_746_EL1809 : EL1809_32157CFD;
	{attribute addProperty Name "Term 747 (EK1110)"}
	{attribute addProperty PreviousPort "Term 746 (EL1809) : B"}
	{attribute addProperty SyncUnit "default"}
	Term_747_EK1110 : EK1110_1FC0878B;
END_STRUCT
END_TYPE

// ---- DUTs/IO/Topology/Term_748_EK1100_BC4343B1.TcDUT
{attribute 'GeneratedUsingTerminal: EK1100-0000-0018'}
{attribute addProperty BoxType "EK1100-0000-0018"}
{attribute addProperty Id "Term_749_EL1809EL1809_32157CFD20Term_750_EL1809EL1809_32157CFD20Term_751_EL1809EL1809_32157CFD20Term_752_EL1809EL1809_32157CFD20Term_753_EL1809EL1809_32157CFD20Term_754_EL1809EL1809_32157CFD20Term_755_EL1809EL1809_32157CFD20Term_756_EL1809EL1809_32157CFD20Term_757_EL1809EL1809_32157CFD20Term_758_EL1809EL1809_32157CFD20Term_759_EL1809EL1809_32157CFD20Term_760_EL1809EL1809_32157CFD20Term_761_EL1809EL1809_32157CFD20Term_762_EL1809EL1809_32157CFD20Term_763_EL1809EL1809_32157CFD20Term_764_EL1809EL1809_32157CFD20Term_765_EL1809EL1809_32157CFD20Term_766_EL1809EL1809_32157CFD20Term_767_EL1809EL1809_32157CFD20Term_768_EL1809EL1809_32157CFD20Term_769_EL1809EL1809_32157CFD20Term_770_EL1809EL1809_32157CFD20Term_771_EL1809EL1809_32157CFD20Term_772_EL1809EL1809_32157CFD20Term_773_EL1809EL1809_32157CFD20Term_774_EL1809EL1809_32157CFD20Term_775_EL1809EL1809_32157CFD20Term_776_EL1809EL1809_32157CFD20Term_777_EL1809EL1809_32157CFD20Term_778_EL1809EL1809_32157CFD20Term_779_EL1809EL1809_32157CFD20Term_780_EL1809EL1809_32157CFD20Term_781_EL1809EL1809_32157CFD20Term_782_EL1809EL1809_32157CFD20Term_783_EL1809EL1809_32157CFD20Term_784_EL1809EL1809_32157CFD20Term_785_EL1809EL1809_32157CFD20Term_786_EL1809EL1809_32157CFD20Term_787_EL1809EL1809_32157CFD20Term_788_EL1809EL1809_32157CFD20Term_789_EL1809EL1809_32157CFD20Term_790_EL1809EL1809_32157CFD20Term_791_EL1809EL1809_32157CFD20Term_792_EL1809EL1809_32157CFD20Term_793_EL1809EL1809_32157CFD20Term_794_EL1809EL1809_32157CFD20Term_795_EL1809EL1809_32157CFD20Term_796_EL1809EL1809_32157CFD20Term_798_EL1809EL1809_32157CFD20Term_799_EL1809EL1809_32157CFD20Term_800_EL1809EL1809_32157CFD20Term_801_EL1809EL1809_32157CFD20Term_802_EL1809EL1809_32157CFD20Term_803_EL1809EL1809_32157CFD20Term_804_EL1809EL1809_32157CFD20Term_805_EL1809EL1809_32157CFD20Term_806_EL1809EL1809_32157CFD20Term_807_EL1809EL1809_32157CFD20Term_808_EL1809EL1809_32157CFD20Term_809_EL1809EL1809_32157CFD20Term_810_EL1809EL1809_32157CFD20Term_811_EL1809EL1809_32157CFD20Term_812_EL1809EL1809_32157CFD20Term_813_EL1809EL1809_32157CFD20Term_814_EL1809EL1809_32157CFD20Term_815_EL1809EL1809_32157CFD20Term_816_EL1809EL1809_32157CFD20Term_817_EL1809EL1809_32157CFD20Term_818_EL1809EL1809_32157CFD20Term_819_EL1809EL1809_32157CFD20Term_820_EL1809EL1809_32157CFD20Term_821_EL1809EL1809_32157CFD20Term_822_EL1809EL1809_32157CFD20Term_823_EL1809EL1809_32157CFD20Term_824_EL1809EL1809_32157CFD20Term_825_EL1809EL1809_32157CFD20Term_826_EL1809EL1809_32157CFD20Term_827_EL1809EL1809_32157CFD20Term_828_EL1809EL1809_32157CFD20Term_859_EL1809EL1809_32157CFD20Term_860_EL1809EL1809_32157CFD20Term_861_EL1809EL1809_32157CFD20Term_862_EL1809EL1809_32157CFD20Term_863_EL1809EL1809_32157CFD20Term_864_EL1809EL1809_32157CFD20Term_865_EL1809EL1809_32157CFD20Term_866_EL1809EL1809_32157CFD20Term_867_EL1809EL1809_32157CFD20Term_868_EL1809EL1809_32157CFD20Term_869_EL1809EL1809_32157CFD20Term_870_EL1809EL1809_32157CFD20Term_871_EL1809EL1809_32157CFD20Term_872_EL1809EL1809_32157CFD20Term_873_EL1809EL1809_32157CFD20Term_874_EL1809EL1809_32157CFD20Term_875_EL1809EL1809_32157CFD20Term_876_EL1809EL1809_32157CFD20Term_877_EL1809EL1809_32157CFD20Term_878_EL1809EL1809_32157CFD20Term_879_EL1809EL1809_32157CFD20Term_880_EK1110EK1110_1FC0878B2"}
{attribute addProperty CRC "3158524849"}
{attribute addProperty Size "2002"}
{attribute addProperty Name "Term 748 (EK1100)"}
TYPE Term_748_EK1100_BC4343B1 EXTENDS EK1100_1FC0878B :
STRUCT
	{attribute addProperty Name "Term 749 (EL1809)"}
	{attribute addProperty PreviousPort "Term 748 (EK1100) : B"}
	{attribute addProperty SyncUnit "default"}
	Term_749_EL1809 : EL1809_32157CFD;
	{attribute addProperty Name "Term 750 (EL1809)"}
	{attribute addProperty PreviousPort "Term 749 (EL1809) : B"}
	{attribute addProperty SyncUnit "default"}
	Term_750_EL1809 : EL1809_32157CFD;
	{attribute addProperty Name "Term 751 (EL1809)"}
	{attribute addProperty PreviousPort "Term 750 (EL1809) : B"}
	{attribute addProperty SyncUnit "default"}
	Term_751_EL1809 : EL1809_32157CFD;
	{attribute addProperty Name "Term 752 (EL1809)"}
	{attribute addProperty PreviousPort "Term 751 (EL1809) : B"}
	{attribute addProperty SyncUnit "default"}
	Term_752_EL1809 : EL1809_32157CFD;
	{attribute addProperty Name "Term 753 (EL1809)"}
	{attribute addProperty PreviousPort "Term 752 (EL1809) : B"}
	{attribute addProperty SyncUnit "default"}
	Term_753_EL1809 : EL1809_32157CFD;
	{attribute addProperty Name "Term 754 (EL1809)"}
	{attribute addProperty PreviousPort "Term 753 (EL1809) : B"}
	{attribute addProperty SyncUnit "default"}
	Term_754_EL1809 : EL1809_32157CFD;
	{attribute addProperty Name "Term 755 (EL1809)"}
	{attribute addProperty PreviousPort "Term 754 (EL1809) : B"}
	{attribute addProperty SyncUnit "default"}
	Term_755_EL1809 : EL1809_32157CFD;
	{attribute addProperty Name "Term 756 (EL1809)"}
	{attribute addProperty PreviousPort "Term 755 (EL1809) : B"}
	{attribute addProperty SyncUnit "default"}
	Term_756_EL1809 : EL1809_32157CFD;
	{attribute addProperty Name "Term 757 (EL1809)"}
	{attribute addProperty PreviousPort "Term 756 (EL1809) : B"}
	{attribute addProperty SyncUnit "default"}
	Term_757_EL1809 : EL1809_32157CFD;
	{attribute addProperty Name "Term 758 (EL1809)"}
	{attribute addProperty PreviousPort "Term 757 (EL1809) : B"}
	{attribute addProperty SyncUnit "default"}
	Term_758_EL1809 : EL1809_32157CFD;
	{attribute addProperty Name "Term 759 (EL1809)"}
	{attribute addProperty PreviousPort "Term 758 (EL1809) : B"}
	{attribute addProperty SyncUnit "default"}
	Term_759_EL1809 : EL1809_32157CFD;
	{attribute addProperty Name "Term 760 (EL1809)"}
	{attribute addProperty PreviousPort "Term 759 (EL1809) : B"}
	{attribute addProperty SyncUnit "default"}
	Term_760_EL1809 : EL1809_32157CFD;
	{attribute addProperty Name "Term 761 (EL1809)"}
	{attribute addProperty PreviousPort "Term 760 (EL1809) : B"}
	{attribute addProperty SyncUnit "default"}
	Term_761_EL1809 : EL1809_32157CFD;
	{attribute addProperty Name "Term 762 (EL1809)"}
	{attribute addProperty PreviousPort "Term 761 (EL1809) : B"}
	{attribute addProperty SyncUnit "default"}
	Term_762_EL1809 : EL1809_32157CFD;
	{attribute addProperty Name "Term 763 (EL1809)"}
	{attribute addProperty PreviousPort "Term 762 (EL1809) : B"}
	{attribute addProperty SyncUnit "default"}
	Term_763_EL1809 : EL1809_32157CFD;
	{attribute addProperty Name "Term 764 (EL1809)"}
	{attribute addProperty PreviousPort "Term 763 (EL1809) : B"}
	{attribute addProperty SyncUnit "default"}
	Term_764_EL1809 : EL1809_32157CFD;
	{attribute addProperty Name "Term 765 (EL1809)"}
	{attribute addProperty PreviousPort "Term 764 (EL1809) : B"}
	{attribute addProperty SyncUnit "default"}
	Term_765_EL1809 : EL1809_32157CFD;
	{attribute addProperty Name "Term 766 (EL1809)"}
	{attribute addProperty PreviousPort "Term 765 (EL1809) : B"}
	{attribute addProperty SyncUnit "default"}
	Term_766_EL1809 : EL1809_32157CFD;
	{attribute addProperty Name "Term 767 (EL1809)"}
	{attribute addProperty PreviousPort "Term 766 (EL1809) : B"}
	{attribute addProperty SyncUnit "default"}
	Term_767_EL1809 : EL1809_32157CFD;
	{attribute addProperty Name "Term 768 (EL1809)"}
	{attribute addProperty PreviousPort "Term 767 (EL1809) : B"}
	{attribute addProperty SyncUnit "default"}
	Term_768_EL1809 : EL1809_32157CFD;
	{attribute addProperty Name "Term 769 (EL1809)"}
	{attribute addProperty PreviousPort "Term 768 (EL1809) : B"}
	{attribute addProperty SyncUnit "default"}
	Term_769_EL1809 : EL1809_32157CFD;
	{attribute addProperty Name "Term 770 (EL1809)"}
	{attribute addProperty PreviousPort "Term 769 (EL1809) : B"}
	{attribute addProperty SyncUnit "default"}
	Term_770_EL1809 : EL1809_32157CFD;
	{attribute addProperty Name "Term 771 (EL1809)"}
	{attribute addProperty PreviousPort "Term 770 (EL1809) : B"}
	{attribute addProperty SyncUnit "default"}
	Term_771_EL1809 : EL1809_32157CFD;
	{attribute addProperty Name "Term 772 (EL1809)"}
	{attribute addProperty PreviousPort "Term 771 (EL1809) : B"}
	{attribute addProperty SyncUnit "default"}
	Term_772_EL1809 : EL1809_32157CFD;
	{attribute addProperty Name "Term 773 (EL1809)"}
	{attribute addProperty PreviousPort "Term 772 (EL1809) : B"}
	{attribute addProperty SyncUnit "default"}
	Term_773_EL1809 : EL1809_32157CFD;
	{attribute addProperty Name "Term 774 (EL1809)"}
	{attribute addProperty PreviousPort "Term 773 (EL1809) : B"}
	{attribute addProperty SyncUnit "default"}
	Term_774_EL1809 : EL1809_32157CFD;
	{attribute addProperty Name "Term 775 (EL1809)"}
	{attribute addProperty PreviousPort "Term 774 (EL1809) : B"}
	{attribute addProperty SyncUnit "default"}
	Term_775_EL1809 : EL1809_32157CFD;
	{attribute addProperty Name "Term 776 (EL1809)"}
	{attribute addProperty PreviousPort "Term 775 (EL1809) : B"}
	{attribute addProperty SyncUnit "default"}
	Term_776_EL1809 : EL1809_32157CFD;
	{attribute addProperty Name "Term 777 (EL1809)"}
	{attribute addProperty PreviousPort "Term 776 (EL1809) : B"}
	{attribute addProperty SyncUnit "default"}
	Term_777_EL1809 : EL1809_32157CFD;
	{attribute addProperty Name "Term 778 (EL1809)"}
	{attribute addProperty PreviousPort "Term 777 (EL1809) : B"}
	{attribute addProperty SyncUnit "default"}
	Term_778_EL1809 : EL1809_32157CFD;
	{attribute addProperty Name "Term 779 (EL1809)"}
	{attribute addProperty PreviousPort "Term 778 (EL1809) : B"}
	{attribute addProperty SyncUnit "default"}
	Term_779_EL1809 : EL1809_32157CFD;
	{attribute addProperty Name "Term 780 (EL1809)"}
	{attribute addProperty PreviousPort "Term 779 (EL1809) : B"}
	{attribute addProperty SyncUnit "default"}
	Term_780_EL1809 : EL1809_32157CFD;
	{attribute addProperty Name "Term 781 (EL1809)"}
	{attribute addProperty PreviousPort "Term 780 (EL1809) : B"}
	{attribute addProperty SyncUnit "default"}
	Term_781_EL1809 : EL1809_32157CFD;
	{attribute addProperty Name "Term 782 (EL1809)"}
	{attribute addProperty PreviousPort "Term 781 (EL1809) : B"}
	{attribute addProperty SyncUnit "default"}
	Term_782_EL1809 : EL1809_32157CFD;
	{attribute addProperty Name "Term 783 (EL1809)"}
	{attribute addProperty PreviousPort "Term 782 (EL1809) : B"}
	{attribute addProperty SyncUnit "default"}
	Term_783_EL1809 : EL1809_32157CFD;
	{attribute addProperty Name "Term 784 (EL1809)"}
	{attribute addProperty PreviousPort "Term 783 (EL1809) : B"}
	{attribute addProperty SyncUnit "default"}
	Term_784_EL1809 : EL1809_32157CFD;
	{attribute addProperty Name "Term 785 (EL1809)"}
	{attribute addProperty PreviousPort "Term 784 (EL1809) : B"}
	{attribute addProperty SyncUnit "default"}
	Term_785_EL1809 : EL1809_32157CFD;
	{attribute addProperty Name "Term 786 (EL1809)"}
	{attribute addProperty PreviousPort "Term 785 (EL1809) : B"}
	{attribute addProperty SyncUnit "default"}
	Term_786_EL1809 : EL1809_32157CFD;
	{attribute addProperty Name "Term 787 (EL1809)"}
	{attribute addProperty PreviousPort "Term 786 (EL1809) : B"}
	{attribute addProperty SyncUnit "default"}
	Term_787_EL1809 : EL1809_32157CFD;
	{attribute addProperty Name "Term 788 (EL1809)"}
	{attribute addProperty PreviousPort "Term 787 (EL1809) : B"}
	{attribute addProperty SyncUnit "default"}
	Term_788_EL1809 : EL1809_32157CFD;
	{attribute addProperty Name "Term 789 (EL1809)"}
	{attribute addProperty PreviousPort "Term 788 (EL1809) : B"}
	{attribute addProperty SyncUnit "default"}
	Term_789_EL1809 : EL1809_32157CFD;
	{attribute addProperty Name "Term 790 (EL1809)"}
	{attribute addProperty PreviousPort "Term 789 (EL1809) : B"}
	{attribute addProperty SyncUnit "default"}
	Term_790_EL1809 : EL1809_32157CFD;
	{attribute addProperty Name "Term 791 (EL1809)"}
	{attribute addProperty PreviousPort "Term 790 (EL1809) : B"}
	{attribute addProperty SyncUnit "default"}
	Term_791_EL1809 : EL1809_32157CFD;
	{attribute addProperty Name "Term 792 (EL1809)"}
	{attribute addProperty PreviousPort "Term 791 (EL1809) : B"}
	{attribute addProperty SyncUnit "default"}
	Term_792_EL1809 : EL1809_32157CFD;
	{attribute addProperty Name "Term 793 (EL1809)"}
	{attribute addProperty PreviousPort "Term 792 (EL1809) : B"}
	{attribute addProperty SyncUnit "default"}
	Term_793_EL1809 : EL1809_32157CFD;
	{attribute addProperty Name "Term 794 (EL1809)"}
	{attribute addProperty PreviousPort "Term 793 (EL1809) : B"}
	{attribute addProperty SyncUnit "default"}
	Term_794_EL1809 : EL1809_32157CFD;
	{attribute addProperty Name "Term 795 (EL1809)"}
	{attribute addProperty PreviousPort "Term 794 (EL1809) : B"}
	{attribute addProperty SyncUnit "default"}
	Term_795_EL1809 : EL1809_32157CFD;
	{attribute addProperty Name "Term 796 (EL1809)"}
	{attribute addProperty PreviousPort "Term 795 (EL1809) : B"}
	{attribute addProperty SyncUnit "default"}
	Term_796_EL1809 : EL1809_32157CFD;
	{attribute addProperty Name "Term 798 (EL1809)"}
	{attribute addProperty PreviousPort "Term 796 (EL1809) : B"}
	{attribute addProperty SyncUnit "default"}
	Term_798_EL1809 : EL1809_32157CFD;
	{attribute addProperty Name "Term 799 (EL1809)"}
	{attribute addProperty PreviousPort "Term 798 (EL1809) : B"}
	{attribute addProperty SyncUnit "default"}
	Term_799_EL1809 : EL1809_32157CFD;
	{attribute addProperty Name "Term 800 (EL1809)"}
	{attribute addProperty PreviousPort "Term 799 (EL1809) : B"}
	{attribute addProperty SyncUnit "default"}
	Term_800_EL1809 : EL1809_32157CFD;
	{attribute addProperty Name "Term 801 (EL1809)"}
	{attribute addProperty PreviousPort "Term 800 (EL1809) : B"}
	{attribute addProperty SyncUnit "default"}
	Term_801_EL1809 : EL1809_32157CFD;
	{attribute addProperty Name "Term 802 (EL1809)"}
	{attribute addProperty PreviousPort "Term 801 (EL1809) : B"}
	{attribute addProperty SyncUnit "default"}
	Term_802_EL1809 : EL1809_32157CFD;
	{attribute addProperty Name "Term 803 (EL1809)"}
	{attribute addProperty PreviousPort "Term 802 (EL1809) : B"}
	{attribute addProperty SyncUnit "default"}
	Term_803_EL1809 : EL1809_32157CFD;
	{attribute addProperty Name "Term 804 (EL1809)"}
	{attribute addProperty PreviousPort "Term 803 (EL1809) : B"}
	{attribute addProperty SyncUnit "default"}
	Term_804_EL1809 : EL1809_32157CFD;
	{attribute addProperty Name "Term 805 (EL1809)"}
	{attribute addProperty PreviousPort "Term 804 (EL1809) : B"}
	{attribute addProperty SyncUnit "default"}
	Term_805_EL1809 : EL1809_32157CFD;
	{attribute addProperty Name "Term 806 (EL1809)"}
	{attribute addProperty PreviousPort "Term 805 (EL1809) : B"}
	{attribute addProperty SyncUnit "default"}
	Term_806_EL1809 : EL1809_32157CFD;
	{attribute addProperty Name "Term 807 (EL1809)"}
	{attribute addProperty PreviousPort "Term 806 (EL1809) : B"}
	{attribute addProperty SyncUnit "default"}
	Term_807_EL1809 : EL1809_32157CFD;
	{attribute addProperty Name "Term 808 (EL1809)"}
	{attribute addProperty PreviousPort "Term 807 (EL1809) : B"}
	{attribute addProperty SyncUnit "default"}
	Term_808_EL1809 : EL1809_32157CFD;
	{attribute addProperty Name "Term 809 (EL1809)"}
	{attribute addProperty PreviousPort "Term 808 (EL1809) : B"}
	{attribute addProperty SyncUnit "default"}
	Term_809_EL1809 : EL1809_32157CFD;
	{attribute addProperty Name "Term 810 (EL1809)"}
	{attribute addProperty PreviousPort "Term 809 (EL1809) : B"}
	{attribute addProperty SyncUnit "default"}
	Term_810_EL1809 : EL1809_32157CFD;
	{attribute addProperty Name "Term 811 (EL1809)"}
	{attribute addProperty PreviousPort "Term 810 (EL1809) : B"}
	{attribute addProperty SyncUnit "default"}
	Term_811_EL1809 : EL1809_32157CFD;
	{attribute addProperty Name "Term 812 (EL1809)"}
	{attribute addProperty PreviousPort "Term 811 (EL1809) : B"}
	{attribute addProperty SyncUnit "default"}
	Term_812_EL1809 : EL1809_32157CFD;
	{attribute addProperty Name "Term 813 (EL1809)"}
	{attribute addProperty PreviousPort "Term 812 (EL1809) : B"}
	{attribute addProperty SyncUnit "default"}
	Term_813_EL1809 : EL1809_32157CFD;
	{attribute addProperty Name "Term 814 (EL1809)"}
	{attribute addProperty PreviousPort "Term 813 (EL1809) : B"}
	{attribute addProperty SyncUnit "default"}
	Term_814_EL1809 : EL1809_32157CFD;
	{attribute addProperty Name "Term 815 (EL1809)"}
	{attribute addProperty PreviousPort "Term 814 (EL1809) : B"}
	{attribute addProperty SyncUnit "default"}
	Term_815_EL1809 : EL1809_32157CFD;
	{attribute addProperty Name "Term 816 (EL1809)"}
	{attribute addProperty PreviousPort "Term 815 (EL1809) : B"}
	{attribute addProperty SyncUnit "default"}
	Term_816_EL1809 : EL1809_32157CFD;
	{attribute addProperty Name "Term 817 (EL1809)"}
	{attribute addProperty PreviousPort "Term 816 (EL1809) : B"}
	{attribute addProperty SyncUnit "default"}
	Term_817_EL1809 : EL1809_32157CFD;
	{attribute addProperty Name "Term 818 (EL1809)"}
	{attribute addProperty PreviousPort "Term 817 (EL1809) : B"}
	{attribute addProperty SyncUnit "default"}
	Term_818_EL1809 : EL1809_32157CFD;
	{attribute addProperty Name "Term 819 (EL1809)"}
	{attribute addProperty PreviousPort "Term 818 (EL1809) : B"}
	{attribute addProperty SyncUnit "default"}
	Term_819_EL1809 : EL1809_32157CFD;
	{attribute addProperty Name "Term 820 (EL1809)"}
	{attribute addProperty PreviousPort "Term 819 (EL1809) : B"}
	{attribute addProperty SyncUnit "default"}
	Term_820_EL1809 : EL1809_32157CFD;
	{attribute addProperty Name "Term 821 (EL1809)"}
	{attribute addProperty PreviousPort "Term 820 (EL1809) : B"}
	{attribute addProperty SyncUnit "default"}
	Term_821_EL1809 : EL1809_32157CFD;
	{attribute addProperty Name "Term 822 (EL1809)"}
	{attribute addProperty PreviousPort "Term 821 (EL1809) : B"}
	{attribute addProperty SyncUnit "default"}
	Term_822_EL1809 : EL1809_32157CFD;
	{attribute addProperty Name "Term 823 (EL1809)"}
	{attribute addProperty PreviousPort "Term 822 (EL1809) : B"}
	{attribute addProperty SyncUnit "default"}
	Term_823_EL1809 : EL1809_32157CFD;
	{attribute addProperty Name "Term 824 (EL1809)"}
	{attribute addProperty PreviousPort "Term 823 (EL1809) : B"}
	{attribute addProperty SyncUnit "default"}
	Term_824_EL1809 : EL1809_32157CFD;
	{attribute addProperty Name "Term 825 (EL1809)"}
	{attribute addProperty PreviousPort "Term 824 (EL1809) : B"}
	{attribute addProperty SyncUnit "default"}
	Term_825_EL1809 : EL1809_32157CFD;
	{attribute addProperty Name "Term 826 (EL1809)"}
	{attribute addProperty PreviousPort "Term 825 (EL1809) : B"}
	{attribute addProperty SyncUnit "default"}
	Term_826_EL1809 : EL1809_32157CFD;
	{attribute addProperty Name "Term 827 (EL1809)"}
	{attribute addProperty PreviousPort "Term 826 (EL1809) : B"}
	{attribute addProperty SyncUnit "default"}
	Term_827_EL1809 : EL1809_32157CFD;
	{attribute addProperty Name "Term 828 (EL1809)"}
	{attribute addProperty PreviousPort "Term 827 (EL1809) : B"}
	{attribute addProperty SyncUnit "default"}
	Term_828_EL1809 : EL1809_32157CFD;
	{attribute addProperty Name "Term 859 (EL1809)"}
	{attribute addProperty PreviousPort "Term 828 (EL1809) : B"}
	{attribute addProperty SyncUnit "default"}
	Term_859_EL1809 : EL1809_32157CFD;
	{attribute addProperty Name "Term 860 (EL1809)"}
	{attribute addProperty PreviousPort "Term 859 (EL1809) : B"}
	{attribute addProperty SyncUnit "default"}
	Term_860_EL1809 : EL1809_32157CFD;
	{attribute addProperty Name "Term 861 (EL1809)"}
	{attribute addProperty PreviousPort "Term 860 (EL1809) : B"}
	{attribute addProperty SyncUnit "default"}
	Term_861_EL1809 : EL1809_32157CFD;
	{attribute addProperty Name "Term 862 (EL1809)"}
	{attribute addProperty PreviousPort "Term 861 (EL1809) : B"}
	{attribute addProperty SyncUnit "default"}
	Term_862_EL1809 : EL1809_32157CFD;
	{attribute addProperty Name "Term 863 (EL1809)"}
	{attribute addProperty PreviousPort "Term 862 (EL1809) : B"}
	{attribute addProperty SyncUnit "default"}
	Term_863_EL1809 : EL1809_32157CFD;
	{attribute addProperty Name "Term 864 (EL1809)"}
	{attribute addProperty PreviousPort "Term 863 (EL1809) : B"}
	{attribute addProperty SyncUnit "default"}
	Term_864_EL1809 : EL1809_32157CFD;
	{attribute addProperty Name "Term 865 (EL1809)"}
	{attribute addProperty PreviousPort "Term 864 (EL1809) : B"}
	{attribute addProperty SyncUnit "default"}
	Term_865_EL1809 : EL1809_32157CFD;
	{attribute addProperty Name "Term 866 (EL1809)"}
	{attribute addProperty PreviousPort "Term 865 (EL1809) : B"}
	{attribute addProperty SyncUnit "default"}
	Term_866_EL1809 : EL1809_32157CFD;
	{attribute addProperty Name "Term 867 (EL1809)"}
	{attribute addProperty PreviousPort "Term 866 (EL1809) : B"}
	{attribute addProperty SyncUnit "default"}
	Term_867_EL1809 : EL1809_32157CFD;
	{attribute addProperty Name "Term 868 (EL1809)"}
	{attribute addProperty PreviousPort "Term 867 (EL1809) : B"}
	{attribute addProperty SyncUnit "default"}
	Term_868_EL1809 : EL1809_32157CFD;
	{attribute addProperty Name "Term 869 (EL1809)"}
	{attribute addProperty PreviousPort "Term 868 (EL1809) : B"}
	{attribute addProperty SyncUnit "default"}
	Term_869_EL1809 : EL1809_32157CFD;
	{attribute addProperty Name "Term 870 (EL1809)"}
	{attribute addProperty PreviousPort "Term 869 (EL1809) : B"}
	{attribute addProperty SyncUnit "default"}
	Term_870_EL1809 : EL1809_32157CFD;
	{attribute addProperty Name "Term 871 (EL1809)"}
	{attribute addProperty PreviousPort "Term 870 (EL1809) : B"}
	{attribute addProperty SyncUnit "default"}
	Term_871_EL1809 : EL1809_32157CFD;
	{attribute addProperty Name "Term 872 (EL1809)"}
	{attribute addProperty PreviousPort "Term 871 (EL1809) : B"}
	{attribute addProperty SyncUnit "default"}
	Term_872_EL1809 : EL1809_32157CFD;
	{attribute addProperty Name "Term 873 (EL1809)"}
	{attribute addProperty PreviousPort "Term 872 (EL1809) : B"}
	{attribute addProperty SyncUnit "default"}
	Term_873_EL1809 : EL1809_32157CFD;
	{attribute addProperty Name "Term 874 (EL1809)"}
	{attribute addProperty PreviousPort "Term 873 (EL1809) : B"}
	{attribute addProperty SyncUnit "default"}
	Term_874_EL1809 : EL1809_32157CFD;
	{attribute addProperty Name "Term 875 (EL1809)"}
	{attribute addProperty PreviousPort "Term 874 (EL1809) : B"}
	{attribute addProperty SyncUnit "default"}
	Term_875_EL1809 : EL1809_32157CFD;
	{attribute addProperty Name "Term 876 (EL1809)"}
	{attribute addProperty PreviousPort "Term 875 (EL1809) : B"}
	{attribute addProperty SyncUnit "default"}
	Term_876_EL1809 : EL1809_32157CFD;
	{attribute addProperty Name "Term 877 (EL1809)"}
	{attribute addProperty PreviousPort "Term 876 (EL1809) : B"}
	{attribute addProperty SyncUnit "default"}
	Term_877_EL1809 : EL1809_32157CFD;
	{attribute addProperty Name "Term 878 (EL1809)"}
	{attribute addProperty PreviousPort "Term 877 (EL1809) : B"}
	{attribute addProperty SyncUnit "default"}
	Term_878_EL1809 : EL1809_32157CFD;
	{attribute addProperty Name "Term 879 (EL1809)"}
	{attribute addProperty PreviousPort "Term 878 (EL1809) : B"}
	{attribute addProperty SyncUnit "default"}
	Term_879_EL1809 : EL1809_32157CFD;
	{attribute addProperty Name "Term 880 (EK1110)"}
	{attribute addProperty PreviousPort "Term 879 (EL1809) : B"}
	{attribute addProperty SyncUnit "default"}
	Term_880_EK1110 : EK1110_1FC0878B;
END_STRUCT
END_TYPE

// ---- DUTs/IO/Topology/Term_881_EK1100_F732F370.TcDUT
{attribute 'GeneratedUsingTerminal: EK1100-0000-0018'}
{attribute addProperty BoxType "EK1100-0000-0018"}
{attribute addProperty Id "Term_882_EL1809EL1809_32157CFD20Term_883_EL1809EL1809_32157CFD20Term_884_EL1809EL1809_32157CFD20Term_885_EL1809EL1809_32157CFD20Term_886_EL1809EL1809_32157CFD20Term_887_EL1809EL1809_32157CFD20Term_888_EL1809EL1809_32157CFD20Term_889_EL1809EL1809_32157CFD20Term_890_EL1809EL1809_32157CFD20Term_891_EL1809EL1809_32157CFD20Term_892_EL1809EL1809_32157CFD20Term_893_EL1809EL1809_32157CFD20Term_894_EL1809EL1809_32157CFD20Term_895_EL1809EL1809_32157CFD20Term_896_EL1809EL1809_32157CFD20Term_897_EL1809EL1809_32157CFD20Term_898_EL1809EL1809_32157CFD20Term_899_EL1809EL1809_32157CFD20Term_900_EL1809EL1809_32157CFD20Term_901_EL1809EL1809_32157CFD20Term_902_EL1809EL1809_32157CFD20Term_903_EL1809EL1809_32157CFD20Term_904_EL1809EL1809_32157CFD20Term_905_EL1809EL1809_32157CFD20Term_906_EL1809EL1809_32157CFD20Term_933_EL1809EL1809_32157CFD20Term_934_EL1809EL1809_32157CFD20Term_935_EL1809EL1809_32157CFD20Term_936_EL1809EL1809_32157CFD20Term_937_EL1809EL1809_32157CFD20Term_938_EL1809EL1809_32157CFD20Term_939_EL1809EL1809_32157CFD20Term_940_EL1809EL1809_32157CFD20Term_941_EL1809EL1809_32157CFD20Term_942_EL1809EL1809_32157CFD20Term_943_EL1809EL1809_32157CFD20Term_944_EL1809EL1809_32157CFD20Term_945_EL1809EL1809_32157CFD20Term_946_EL1809EL1809_32157CFD20Term_947_EL1809EL1809_32157CFD20Term_948_EL1809EL1809_32157CFD20Term_949_EL1809EL1809_32157CFD20Term_950_EL1809EL1809_32157CFD20Term_951_EL1809EL1809_32157CFD20Term_952_EL1809EL1809_32157CFD20Term_953_EL1809EL1809_32157CFD20Term_954_EL1809EL1809_32157CFD20Term_955_EL1809EL1809_32157CFD20Term_956_EL1809EL1809_32157CFD20Term_957_EL1809EL1809_32157CFD20Term_958_EL1809EL1809_32157CFD20Term_959_EL1809EL1809_32157CFD20Term_960_EL1809EL1809_32157CFD20Term_961_EL1809EL1809_32157CFD20Term_962_EL1809EL1809_32157CFD20Term_963_EL1809EL1809_32157CFD20Term_964_EL1809EL1809_32157CFD20Term_965_EL1809EL1809_32157CFD20Term_967_EL1809EL1809_32157CFD20Term_968_EL1809EL1809_32157CFD20Term_969_EL1809EL1809_32157CFD20Term_970_EL1809EL1809_32157CFD20Term_971_EL1809EL1809_32157CFD20Term_972_EL1809EL1809_32157CFD20Term_973_EL1809EL1809_32157CFD20Term_974_EL1809EL1809_32157CFD20Term_975_EL1809EL1809_32157CFD20Term_976_EL1809EL1809_32157CFD20Term_977_EL1809EL1809_32157CFD20Term_978_EL1809EL1809_32157CFD20Term_979_EL1809EL1809_32157CFD20Term_980_EL1809EL1809_32157CFD20Term_981_EL1809EL1809_32157CFD20Term_982_EL1809EL1809_32157CFD20Term_983_EL1809EL1809_32157CFD20Term_984_EL1809EL1809_32157CFD20Term_986_EL1809EL1809_32157CFD20Term_987_EL1809EL1809_32157CFD20Term_988_EL1809EL1809_32157CFD20Term_989_EL1809EL1809_32157CFD20Term_1025_EL1809EL1809_32157CFD20Term_1026_EL1809EL1809_32157CFD20Term_1027_EL1809EL1809_32157CFD20Term_1028_EL1809EL1809_32157CFD20Term_1029_EL1809EL1809_32157CFD20Term_1030_EL1809EL1809_32157CFD20Term_1031_EL1809EL1809_32157CFD20Term_1032_EL1809EL1809_32157CFD20Term_1033_EL1809EL1809_32157CFD20Term_1034_EL1809EL1809_32157CFD20Term_1035_EL1809EL1809_32157CFD20Term_1036_EL1809EL1809_32157CFD20Term_1038_EL1809EL1809_32157CFD20Term_1039_EL1809EL1809_32157CFD20Term_1040_EL1809EL1809_32157CFD20Term_1041_EL1809EL1809_32157CFD20Term_1042_EL1809EL1809_32157CFD20Term_1043_EL1809EL1809_32157CFD20Term_1044_EL1809EL1809_32157CFD20Term_1045_EL1809EL1809_32157CFD20Term_1046_EK1110EK1110_1FC0878B2"}
{attribute addProperty CRC "4147311472"}
{attribute addProperty Size "2002"}
{attribute addProperty Name "Term 881 (EK1100)"}
TYPE Term_881_EK1100_F732F370 EXTENDS EK1100_1FC0878B :
STRUCT
	{attribute addProperty Name "Term 882 (EL1809)"}
	{attribute addProperty PreviousPort "Term 881 (EK1100) : B"}
	{attribute addProperty SyncUnit "default"}
	Term_882_EL1809 : EL1809_32157CFD;
	{attribute addProperty Name "Term 883 (EL1809)"}
	{attribute addProperty PreviousPort "Term 882 (EL1809) : B"}
	{attribute addProperty SyncUnit "default"}
	Term_883_EL1809 : EL1809_32157CFD;
	{attribute addProperty Name "Term 884 (EL1809)"}
	{attribute addProperty PreviousPort "Term 883 (EL1809) : B"}
	{attribute addProperty SyncUnit "default"}
	Term_884_EL1809 : EL1809_32157CFD;
	{attribute addProperty Name "Term 885 (EL1809)"}
	{attribute addProperty PreviousPort "Term 884 (EL1809) : B"}
	{attribute addProperty SyncUnit "default"}
	Term_885_EL1809 : EL1809_32157CFD;
	{attribute addProperty Name "Term 886 (EL1809)"}
	{attribute addProperty PreviousPort "Term 885 (EL1809) : B"}
	{attribute addProperty SyncUnit "default"}
	Term_886_EL1809 : EL1809_32157CFD;
	{attribute addProperty Name "Term 887 (EL1809)"}
	{attribute addProperty PreviousPort "Term 886 (EL1809) : B"}
	{attribute addProperty SyncUnit "default"}
	Term_887_EL1809 : EL1809_32157CFD;
	{attribute addProperty Name "Term 888 (EL1809)"}
	{attribute addProperty PreviousPort "Term 887 (EL1809) : B"}
	{attribute addProperty SyncUnit "default"}
	Term_888_EL1809 : EL1809_32157CFD;
	{attribute addProperty Name "Term 889 (EL1809)"}
	{attribute addProperty PreviousPort "Term 888 (EL1809) : B"}
	{attribute addProperty SyncUnit "default"}
	Term_889_EL1809 : EL1809_32157CFD;
	{attribute addProperty Name "Term 890 (EL1809)"}
	{attribute addProperty PreviousPort "Term 889 (EL1809) : B"}
	{attribute addProperty SyncUnit "default"}
	Term_890_EL1809 : EL1809_32157CFD;
	{attribute addProperty Name "Term 891 (EL1809)"}
	{attribute addProperty PreviousPort "Term 890 (EL1809) : B"}
	{attribute addProperty SyncUnit "default"}
	Term_891_EL1809 : EL1809_32157CFD;
	{attribute addProperty Name "Term 892 (EL1809)"}
	{attribute addProperty PreviousPort "Term 891 (EL1809) : B"}
	{attribute addProperty SyncUnit "default"}
	Term_892_EL1809 : EL1809_32157CFD;
	{attribute addProperty Name "Term 893 (EL1809)"}
	{attribute addProperty PreviousPort "Term 892 (EL1809) : B"}
	{attribute addProperty SyncUnit "default"}
	Term_893_EL1809 : EL1809_32157CFD;
	{attribute addProperty Name "Term 894 (EL1809)"}
	{attribute addProperty PreviousPort "Term 893 (EL1809) : B"}
	{attribute addProperty SyncUnit "default"}
	Term_894_EL1809 : EL1809_32157CFD;
	{attribute addProperty Name "Term 895 (EL1809)"}
	{attribute addProperty PreviousPort "Term 894 (EL1809) : B"}
	{attribute addProperty SyncUnit "default"}
	Term_895_EL1809 : EL1809_32157CFD;
	{attribute addProperty Name "Term 896 (EL1809)"}
	{attribute addProperty PreviousPort "Term 895 (EL1809) : B"}
	{attribute addProperty SyncUnit "default"}
	Term_896_EL1809 : EL1809_32157CFD;
	{attribute addProperty Name "Term 897 (EL1809)"}
	{attribute addProperty PreviousPort "Term 896 (EL1809) : B"}
	{attribute addProperty SyncUnit "default"}
	Term_897_EL1809 : EL1809_32157CFD;
	{attribute addProperty Name "Term 898 (EL1809)"}
	{attribute addProperty PreviousPort "Term 897 (EL1809) : B"}
	{attribute addProperty SyncUnit "default"}
	Term_898_EL1809 : EL1809_32157CFD;
	{attribute addProperty Name "Term 899 (EL1809)"}
	{attribute addProperty PreviousPort "Term 898 (EL1809) : B"}
	{attribute addProperty SyncUnit "default"}
	Term_899_EL1809 : EL1809_32157CFD;
	{attribute addProperty Name "Term 900 (EL1809)"}
	{attribute addProperty PreviousPort "Term 899 (EL1809) : B"}
	{attribute addProperty SyncUnit "default"}
	Term_900_EL1809 : EL1809_32157CFD;
	{attribute addProperty Name "Term 901 (EL1809)"}
	{attribute addProperty PreviousPort "Term 900 (EL1809) : B"}
	{attribute addProperty SyncUnit "default"}
	Term_901_EL1809 : EL1809_32157CFD;
	{attribute addProperty Name "Term 902 (EL1809)"}
	{attribute addProperty PreviousPort "Term 901 (EL1809) : B"}
	{attribute addProperty SyncUnit "default"}
	Term_902_EL1809 : EL1809_32157CFD;
	{attribute addProperty Name "Term 903 (EL1809)"}
	{attribute addProperty PreviousPort "Term 902 (EL1809) : B"}
	{attribute addProperty SyncUnit "default"}
	Term_903_EL1809 : EL1809_32157CFD;
	{attribute addProperty Name "Term 904 (EL1809)"}
	{attribute addProperty PreviousPort "Term 903 (EL1809) : B"}
	{attribute addProperty SyncUnit "default"}
	Term_904_EL1809 : EL1809_32157CFD;
	{attribute addProperty Name "Term 905 (EL1809)"}
	{attribute addProperty PreviousPort "Term 904 (EL1809) : B"}
	{attribute addProperty SyncUnit "default"}
	Term_905_EL1809 : EL1809_32157CFD;
	{attribute addProperty Name "Term 906 (EL1809)"}
	{attribute addProperty PreviousPort "Term 905 (EL1809) : B"}
	{attribute addProperty SyncUnit "default"}
	Term_906_EL1809 : EL1809_32157CFD;
	{attribute addProperty Name "Term 933 (EL1809)"}
	{attribute addProperty PreviousPort "Term 906 (EL1809) : B"}
	{attribute addProperty SyncUnit "default"}
	Term_933_EL1809 : EL1809_32157CFD;
	{attribute addProperty Name "Term 934 (EL1809)"}
	{attribute addProperty PreviousPort "Term 933 (EL1809) : B"}
	{attribute addProperty SyncUnit "default"}
	Term_934_EL1809 : EL1809_32157CFD;
	{attribute addProperty Name "Term 935 (EL1809)"}
	{attribute addProperty PreviousPort "Term 934 (EL1809) : B"}
	{attribute addProperty SyncUnit "default"}
	Term_935_EL1809 : EL1809_32157CFD;
	{attribute addProperty Name "Term 936 (EL1809)"}
	{attribute addProperty PreviousPort "Term 935 (EL1809) : B"}
	{attribute addProperty SyncUnit "default"}
	Term_936_EL1809 : EL1809_32157CFD;
	{attribute addProperty Name "Term 937 (EL1809)"}
	{attribute addProperty PreviousPort "Term 936 (EL1809) : B"}
	{attribute addProperty SyncUnit "default"}
	Term_937_EL1809 : EL1809_32157CFD;
	{attribute addProperty Name "Term 938 (EL1809)"}
	{attribute addProperty PreviousPort "Term 937 (EL1809) : B"}
	{attribute addProperty SyncUnit "default"}
	Term_938_EL1809 : EL1809_32157CFD;
	{attribute addProperty Name "Term 939 (EL1809)"}
	{attribute addProperty PreviousPort "Term 938 (EL1809) : B"}
	{attribute addProperty SyncUnit "default"}
	Term_939_EL1809 : EL1809_32157CFD;
	{attribute addProperty Name "Term 940 (EL1809)"}
	{attribute addProperty PreviousPort "Term 939 (EL1809) : B"}
	{attribute addProperty SyncUnit "default"}
	Term_940_EL1809 : EL1809_32157CFD;
	{attribute addProperty Name "Term 941 (EL1809)"}
	{attribute addProperty PreviousPort "Term 940 (EL1809) : B"}
	{attribute addProperty SyncUnit "default"}
	Term_941_EL1809 : EL1809_32157CFD;
	{attribute addProperty Name "Term 942 (EL1809)"}
	{attribute addProperty PreviousPort "Term 941 (EL1809) : B"}
	{attribute addProperty SyncUnit "default"}
	Term_942_EL1809 : EL1809_32157CFD;
	{attribute addProperty Name "Term 943 (EL1809)"}
	{attribute addProperty PreviousPort "Term 942 (EL1809) : B"}
	{attribute addProperty SyncUnit "default"}
	Term_943_EL1809 : EL1809_32157CFD;
	{attribute addProperty Name "Term 944 (EL1809)"}
	{attribute addProperty PreviousPort "Term 943 (EL1809) : B"}
	{attribute addProperty SyncUnit "default"}
	Term_944_EL1809 : EL1809_32157CFD;
	{attribute addProperty Name "Term 945 (EL1809)"}
	{attribute addProperty PreviousPort "Term 944 (EL1809) : B"}
	{attribute addProperty SyncUnit "default"}
	Term_945_EL1809 : EL1809_32157CFD;
	{attribute addProperty Name "Term 946 (EL1809)"}
	{attribute addProperty PreviousPort "Term 945 (EL1809) : B"}
	{attribute addProperty SyncUnit "default"}
	Term_946_EL1809 : EL1809_32157CFD;
	{attribute addProperty Name "Term 947 (EL1809)"}
	{attribute addProperty PreviousPort "Term 946 (EL1809) : B"}
	{attribute addProperty SyncUnit "default"}
	Term_947_EL1809 : EL1809_32157CFD;
	{attribute addProperty Name "Term 948 (EL1809)"}
	{attribute addProperty PreviousPort "Term 947 (EL1809) : B"}
	{attribute addProperty SyncUnit "default"}
	Term_948_EL1809 : EL1809_32157CFD;
	{attribute addProperty Name "Term 949 (EL1809)"}
	{attribute addProperty PreviousPort "Term 948 (EL1809) : B"}
	{attribute addProperty SyncUnit "default"}
	Term_949_EL1809 : EL1809_32157CFD;
	{attribute addProperty Name "Term 950 (EL1809)"}
	{attribute addProperty PreviousPort "Term 949 (EL1809) : B"}
	{attribute addProperty SyncUnit "default"}
	Term_950_EL1809 : EL1809_32157CFD;
	{attribute addProperty Name "Term 951 (EL1809)"}
	{attribute addProperty PreviousPort "Term 950 (EL1809) : B"}
	{attribute addProperty SyncUnit "default"}
	Term_951_EL1809 : EL1809_32157CFD;
	{attribute addProperty Name "Term 952 (EL1809)"}
	{attribute addProperty PreviousPort "Term 951 (EL1809) : B"}
	{attribute addProperty SyncUnit "default"}
	Term_952_EL1809 : EL1809_32157CFD;
	{attribute addProperty Name "Term 953 (EL1809)"}
	{attribute addProperty PreviousPort "Term 952 (EL1809) : B"}
	{attribute addProperty SyncUnit "default"}
	Term_953_EL1809 : EL1809_32157CFD;
	{attribute addProperty Name "Term 954 (EL1809)"}
	{attribute addProperty PreviousPort "Term 953 (EL1809) : B"}
	{attribute addProperty SyncUnit "default"}
	Term_954_EL1809 : EL1809_32157CFD;
	{attribute addProperty Name "Term 955 (EL1809)"}
	{attribute addProperty PreviousPort "Term 954 (EL1809) : B"}
	{attribute addProperty SyncUnit "default"}
	Term_955_EL1809 : EL1809_32157CFD;
	{attribute addProperty Name "Term 956 (EL1809)"}
	{attribute addProperty PreviousPort "Term 955 (EL1809) : B"}
	{attribute addProperty SyncUnit "default"}
	Term_956_EL1809 : EL1809_32157CFD;
	{attribute addProperty Name "Term 957 (EL1809)"}
	{attribute addProperty PreviousPort "Term 956 (EL1809) : B"}
	{attribute addProperty SyncUnit "default"}
	Term_957_EL1809 : EL1809_32157CFD;
	{attribute addProperty Name "Term 958 (EL1809)"}
	{attribute addProperty PreviousPort "Term 957 (EL1809) : B"}
	{attribute addProperty SyncUnit "default"}
	Term_958_EL1809 : EL1809_32157CFD;
	{attribute addProperty Name "Term 959 (EL1809)"}
	{attribute addProperty PreviousPort "Term 958 (EL1809) : B"}
	{attribute addProperty SyncUnit "default"}
	Term_959_EL1809 : EL1809_32157CFD;
	{attribute addProperty Name "Term 960 (EL1809)"}
	{attribute addProperty PreviousPort "Term 959 (EL1809) : B"}
	{attribute addProperty SyncUnit "default"}
	Term_960_EL1809 : EL1809_32157CFD;
	{attribute addProperty Name "Term 961 (EL1809)"}
	{attribute addProperty PreviousPort "Term 960 (EL1809) : B"}
	{attribute addProperty SyncUnit "default"}
	Term_961_EL1809 : EL1809_32157CFD;
	{attribute addProperty Name "Term 962 (EL1809)"}
	{attribute addProperty PreviousPort "Term 961 (EL1809) : B"}
	{attribute addProperty SyncUnit "default"}
	Term_962_EL1809 : EL1809_32157CFD;
	{attribute addProperty Name "Term 963 (EL1809)"}
	{attribute addProperty PreviousPort "Term 962 (EL1809) : B"}
	{attribute addProperty SyncUnit "default"}
	Term_963_EL1809 : EL1809_32157CFD;
	{attribute addProperty Name "Term 964 (EL1809)"}
	{attribute addProperty PreviousPort "Term 963 (EL1809) : B"}
	{attribute addProperty SyncUnit "default"}
	Term_964_EL1809 : EL1809_32157CFD;
	{attribute addProperty Name "Term 965 (EL1809)"}
	{attribute addProperty PreviousPort "Term 964 (EL1809) : B"}
	{attribute addProperty SyncUnit "default"}
	Term_965_EL1809 : EL1809_32157CFD;
	{attribute addProperty Name "Term 967 (EL1809)"}
	{attribute addProperty PreviousPort "Term 965 (EL1809) : B"}
	{attribute addProperty SyncUnit "default"}
	Term_967_EL1809 : EL1809_32157CFD;
	{attribute addProperty Name "Term 968 (EL1809)"}
	{attribute addProperty PreviousPort "Term 967 (EL1809) : B"}
	{attribute addProperty SyncUnit "default"}
	Term_968_EL1809 : EL1809_32157CFD;
	{attribute addProperty Name "Term 969 (EL1809)"}
	{attribute addProperty PreviousPort "Term 968 (EL1809) : B"}
	{attribute addProperty SyncUnit "default"}
	Term_969_EL1809 : EL1809_32157CFD;
	{attribute addProperty Name "Term 970 (EL1809)"}
	{attribute addProperty PreviousPort "Term 969 (EL1809) : B"}
	{attribute addProperty SyncUnit "default"}
	Term_970_EL1809 : EL1809_32157CFD;
	{attribute addProperty Name "Term 971 (EL1809)"}
	{attribute addProperty PreviousPort "Term 970 (EL1809) : B"}
	{attribute addProperty SyncUnit "default"}
	Term_971_EL1809 : EL1809_32157CFD;
	{attribute addProperty Name "Term 972 (EL1809)"}
	{attribute addProperty PreviousPort "Term 971 (EL1809) : B"}
	{attribute addProperty SyncUnit "default"}
	Term_972_EL1809 : EL1809_32157CFD;
	{attribute addProperty Name "Term 973 (EL1809)"}
	{attribute addProperty PreviousPort "Term 972 (EL1809) : B"}
	{attribute addProperty SyncUnit "default"}
	Term_973_EL1809 : EL1809_32157CFD;
	{attribute addProperty Name "Term 974 (EL1809)"}
	{attribute addProperty PreviousPort "Term 973 (EL1809) : B"}
	{attribute addProperty SyncUnit "default"}
	Term_974_EL1809 : EL1809_32157CFD;
	{attribute addProperty Name "Term 975 (EL1809)"}
	{attribute addProperty PreviousPort "Term 974 (EL1809) : B"}
	{attribute addProperty SyncUnit "default"}
	Term_975_EL1809 : EL1809_32157CFD;
	{attribute addProperty Name "Term 976 (EL1809)"}
	{attribute addProperty PreviousPort "Term 975 (EL1809) : B"}
	{attribute addProperty SyncUnit "default"}
	Term_976_EL1809 : EL1809_32157CFD;
	{attribute addProperty Name "Term 977 (EL1809)"}
	{attribute addProperty PreviousPort "Term 976 (EL1809) : B"}
	{attribute addProperty SyncUnit "default"}
	Term_977_EL1809 : EL1809_32157CFD;
	{attribute addProperty Name "Term 978 (EL1809)"}
	{attribute addProperty PreviousPort "Term 977 (EL1809) : B"}
	{attribute addProperty SyncUnit "default"}
	Term_978_EL1809 : EL1809_32157CFD;
	{attribute addProperty Name "Term 979 (EL1809)"}
	{attribute addProperty PreviousPort "Term 978 (EL1809) : B"}
	{attribute addProperty SyncUnit "default"}
	Term_979_EL1809 : EL1809_32157CFD;
	{attribute addProperty Name "Term 980 (EL1809)"}
	{attribute addProperty PreviousPort "Term 979 (EL1809) : B"}
	{attribute addProperty SyncUnit "default"}
	Term_980_EL1809 : EL1809_32157CFD;
	{attribute addProperty Name "Term 981 (EL1809)"}
	{attribute addProperty PreviousPort "Term 980 (EL1809) : B"}
	{attribute addProperty SyncUnit "default"}
	Term_981_EL1809 : EL1809_32157CFD;
	{attribute addProperty Name "Term 982 (EL1809)"}
	{attribute addProperty PreviousPort "Term 981 (EL1809) : B"}
	{attribute addProperty SyncUnit "default"}
	Term_982_EL1809 : EL1809_32157CFD;
	{attribute addProperty Name "Term 983 (EL1809)"}
	{attribute addProperty PreviousPort "Term 982 (EL1809) : B"}
	{attribute addProperty SyncUnit "default"}
	Term_983_EL1809 : EL1809_32157CFD;
	{attribute addProperty Name "Term 984 (EL1809)"}
	{attribute addProperty PreviousPort "Term 983 (EL1809) : B"}
	{attribute addProperty SyncUnit "default"}
	Term_984_EL1809 : EL1809_32157CFD;
	{attribute addProperty Name "Term 986 (EL1809)"}
	{attribute addProperty PreviousPort "Term 984 (EL1809) : B"}
	{attribute addProperty SyncUnit "default"}
	Term_986_EL1809 : EL1809_32157CFD;
	{attribute addProperty Name "Term 987 (EL1809)"}
	{attribute addProperty PreviousPort "Term 986 (EL1809) : B"}
	{attribute addProperty SyncUnit "default"}
	Term_987_EL1809 : EL1809_32157CFD;
	{attribute addProperty Name "Term 988 (EL1809)"}
	{attribute addProperty PreviousPort "Term 987 (EL1809) : B"}
	{attribute addProperty SyncUnit "default"}
	Term_988_EL1809 : EL1809_32157CFD;
	{attribute addProperty Name "Term 989 (EL1809)"}
	{attribute addProperty PreviousPort "Term 988 (EL1809) : B"}
	{attribute addProperty SyncUnit "default"}
	Term_989_EL1809 : EL1809_32157CFD;
	{attribute addProperty Name "Term 1025 (EL1809)"}
	{attribute addProperty PreviousPort "Term 989 (EL1809) : B"}
	{attribute addProperty SyncUnit "default"}
	Term_1025_EL1809 : EL1809_32157CFD;
	{attribute addProperty Name "Term 1026 (EL1809)"}
	{attribute addProperty PreviousPort "Term 1025 (EL1809) : B"}
	{attribute addProperty SyncUnit "default"}
	Term_1026_EL1809 : EL1809_32157CFD;
	{attribute addProperty Name "Term 1027 (EL1809)"}
	{attribute addProperty PreviousPort "Term 1026 (EL1809) : B"}
	{attribute addProperty SyncUnit "default"}
	Term_1027_EL1809 : EL1809_32157CFD;
	{attribute addProperty Name "Term 1028 (EL1809)"}
	{attribute addProperty PreviousPort "Term 1027 (EL1809) : B"}
	{attribute addProperty SyncUnit "default"}
	Term_1028_EL1809 : EL1809_32157CFD;
	{attribute addProperty Name "Term 1029 (EL1809)"}
	{attribute addProperty PreviousPort "Term 1028 (EL1809) : B"}
	{attribute addProperty SyncUnit "default"}
	Term_1029_EL1809 : EL1809_32157CFD;
	{attribute addProperty Name "Term 1030 (EL1809)"}
	{attribute addProperty PreviousPort "Term 1029 (EL1809) : B"}
	{attribute addProperty SyncUnit "default"}
	Term_1030_EL1809 : EL1809_32157CFD;
	{attribute addProperty Name "Term 1031 (EL1809)"}
	{attribute addProperty PreviousPort "Term 1030 (EL1809) : B"}
	{attribute addProperty SyncUnit "default"}
	Term_1031_EL1809 : EL1809_32157CFD;
	{attribute addProperty Name "Term 1032 (EL1809)"}
	{attribute addProperty PreviousPort "Term 1031 (EL1809) : B"}
	{attribute addProperty SyncUnit "default"}
	Term_1032_EL1809 : EL1809_32157CFD;
	{attribute addProperty Name "Term 1033 (EL1809)"}
	{attribute addProperty PreviousPort "Term 1032 (EL1809) : B"}
	{attribute addProperty SyncUnit "default"}
	Term_1033_EL1809 : EL1809_32157CFD;
	{attribute addProperty Name "Term 1034 (EL1809)"}
	{attribute addProperty PreviousPort "Term 1033 (EL1809) : B"}
	{attribute addProperty SyncUnit "default"}
	Term_1034_EL1809 : EL1809_32157CFD;
	{attribute addProperty Name "Term 1035 (EL1809)"}
	{attribute addProperty PreviousPort "Term 1034 (EL1809) : B"}
	{attribute addProperty SyncUnit "default"}
	Term_1035_EL1809 : EL1809_32157CFD;
	{attribute addProperty Name "Term 1036 (EL1809)"}
	{attribute addProperty PreviousPort "Term 1035 (EL1809) : B"}
	{attribute addProperty SyncUnit "default"}
	Term_1036_EL1809 : EL1809_32157CFD;
	{attribute addProperty Name "Term 1038 (EL1809)"}
	{attribute addProperty PreviousPort "Term 1036 (EL1809) : B"}
	{attribute addProperty SyncUnit "default"}
	Term_1038_EL1809 : EL1809_32157CFD;
	{attribute addProperty Name "Term 1039 (EL1809)"}
	{attribute addProperty PreviousPort "Term 1038 (EL1809) : B"}
	{attribute addProperty SyncUnit "default"}
	Term_1039_EL1809 : EL1809_32157CFD;
	{attribute addProperty Name "Term 1040 (EL1809)"}
	{attribute addProperty PreviousPort "Term 1039 (EL1809) : B"}
	{attribute addProperty SyncUnit "default"}
	Term_1040_EL1809 : EL1809_32157CFD;
	{attribute addProperty Name "Term 1041 (EL1809)"}
	{attribute addProperty PreviousPort "Term 1040 (EL1809) : B"}
	{attribute addProperty SyncUnit "default"}
	Term_1041_EL1809 : EL1809_32157CFD;
	{attribute addProperty Name "Term 1042 (EL1809)"}
	{attribute addProperty PreviousPort "Term 1041 (EL1809) : B"}
	{attribute addProperty SyncUnit "default"}
	Term_1042_EL1809 : EL1809_32157CFD;
	{attribute addProperty Name "Term 1043 (EL1809)"}
	{attribute addProperty PreviousPort "Term 1042 (EL1809) : B"}
	{attribute addProperty SyncUnit "default"}
	Term_1043_EL1809 : EL1809_32157CFD;
	{attribute addProperty Name "Term 1044 (EL1809)"}
	{attribute addProperty PreviousPort "Term 1043 (EL1809) : B"}
	{attribute addProperty SyncUnit "default"}
	Term_1044_EL1809 : EL1809_32157CFD;
	{attribute addProperty Name "Term 1045 (EL1809)"}
	{attribute addProperty PreviousPort "Term 1044 (EL1809) : B"}
	{attribute addProperty SyncUnit "default"}
	Term_1045_EL1809 : EL1809_32157CFD;
	{attribute addProperty Name "Term 1046 (EK1110)"}
	{attribute addProperty PreviousPort "Term 1045 (EL1809) : B"}
	{attribute addProperty SyncUnit "default"}
	Term_1046_EK1110 : EK1110_1FC0878B;
END_STRUCT
END_TYPE

